(* IEC 61131-3 sources: Test-Git_ESME26/TestProgettoESME_26.fbsproj/AxisModuleLib Migration/DiagSource/AXM_FB_AxisModuleDiagSource.fb.st^, 38 files *)

(* ---- CancelWriting.meth.st ---- *)
{attribute 'conditionalshow_all_locals'}
METHOD INTERNAL CancelWriting : BOOL
VAR_INPUT
END_VAR

(* Deactivate writing if we are (for whatever reason) no longer adressed.
   May happen in case network connection with Diagnostics is disrupted or Source will be disabled *)

THIS^.diOldCmd			:= 0;
THIS^.diCmdExecState	:= 0;

(* ---- DiagQuit.meth.st ---- *)
{attribute 'conditionalshow_all_locals'}
METHOD INTERNAL DiagQuit : BOOL
VAR_INPUT
END_VAR

IF THIS^.i_xEnable AND THIS^.q_xActive AND THIS^.q_etDiag <> GD.ET_Diag.Ok AND THIS^.diState = 0 THEN

	THIS^.rtrigDiagQuit(CLK := THIS^.i_xDiagQuit);
	IF THIS^.rtrigDiagQuit.Q THEN
		CancelWriting();

		THIS^.udiOwnSourceId	:= 0;

		THIS^.fbTreeWriter.FB_Init(bInitRetains := FALSE, bInCopyCode := FALSE);

		THIS^.q_xReady		:= TRUE;
		THIS^.q_etDiag		:= GD.ET_Diag.Ok;
		THIS^.q_etDiagExt	:= AXM_ET_DiagExt.WaitUntilDiagnosticsManagerReady;
		THIS^.q_sMsg		:= '';

		THIS^.diState := 10;
	END_IF

END_IF

(* ---- ExceptionDuringWriting.meth.st ---- *)
{attribute 'conditionalshow_all_locals'}
METHOD INTERNAL ExceptionDuringWriting : BOOL
VAR_INPUT
END_VAR

(* exception during writing *)
CASE THIS^.etDiagExtTPL OF
	TPL.ET_DiagExt.TreeStartAlreadySuccessfullyCalled,
	TPL.ET_DiagExt.FileIdNotSet,
	TPL.ET_DiagExt.FileIdInvalid,
	TPL.ET_DiagExt.FileNotOpen,
	TPL.ET_DiagExt.UnexpectedFeedback,
	TPL.ET_DiagExt.TreeStartNotCalled,
	TPL.ET_DiagExt.TreeStartNotSuccessfullyCalled,
	TPL.ET_DiagExt.NoMoreNodeOpen,
	TPL.ET_DiagExt.CallTreeStartFirst,
	TPL.ET_DiagExt.NodesStillOpen:

		SetDiagOutputs(	i_etDiag	:= GD.ET_Diag.UnexpectedProgramBehavior,
						i_etDiagExt	:= AXM_ET_DiagExt.UnexpectedFeedback,
						i_sMsg		:= SE_CTBX.FC_MultiConcat(	i_sString1	:= 'FB_TreeWriter: ',
																i_sString2	:= GD.FC_EtDiagToString(THIS^.etDiag),
																i_sString3	:= ' - ',
																i_sString4	:= TPL.FC_EtDiagExtToString(THIS^.etDiagExtTPL)
															 )
					  );
	ELSE
		SetDiagOutputs(	i_etDiag	:= GD.ET_Diag.UnexpectedProgramBehavior,
						i_etDiagExt	:= AXM_ET_DiagExt.UnexpectedFeedback,
						i_sMsg		:= SE_CTBX.FC_MultiConcat(	i_sString1	:= 'FB_TreeWriter: ',
																i_sString2	:= GD.FC_EtDiagToString(THIS^.etDiag),
																i_sString3	:= ' - ',
																i_sString4	:= TPL.FC_EtDiagExtToString(THIS^.etDiagExtTPL)
															  )
					   );
END_CASE

CancelWriting();

(* ---- SetDiagOutputs.meth.st ---- *)
{attribute 'conditionalshow_all_locals'}
METHOD INTERNAL SetDiagOutputs : BOOL
VAR_INPUT
	i_etDiag		: GD.ET_Diag;
	i_etDiagExt		: AXM_ET_DiagExt;
	i_sMsg			: STRING[80];
END_VAR

IF THIS^.q_etDiag = GD.ET_Diag.Ok OR i_etDiagExt = AXM_ET_DiagExt.Disabled THEN

	IF i_etDiag <> GD.ET_Diag.Ok OR i_etDiagExt = AXM_ET_DiagExt.Disabled THEN

		IF i_etDiag <> GD.ET_Diag.Ok THEN
			THIS^.iq_stComStructure.iq_diCmd := -THIS^.iq_stComStructure.iq_diCmd;
		END_IF

		IF i_etDiagExt = AXM_ET_DiagExt.Disabled THEN
			THIS^.q_xActive := FALSE;

			CancelWriting();
		END_IF

		THIS^.q_xReady := FALSE;
		THIS^.diState := 0;
	END_IF

	THIS^.q_etDiag		:= i_etDiag;
	THIS^.q_etDiagExt	:= i_etDiagExt;
	THIS^.q_sMsg		:= i_sMsg;

END_IF

(* ---- WriteDiagDataControl.meth.st ---- *)
{attribute 'conditionalshow_all_locals'}
METHOD INTERNAL WriteDiagDataControl : BOOL
VAR_INPUT
END_VAR

IF (THIS^.diOldCmd <> THIS^.iq_stComStructure.iq_diCmd AND THIS^.iq_stComStructure.iq_diCmd > 0) THEN

	THIS^.diOldCmd := THIS^.iq_stComStructure.iq_diCmd;

	(* new command, start execution *)
	CASE THIS^.iq_stComStructure.iq_diCmd OF

		1: (* write diag data to file *)
			IF (THIS^.iq_stComStructure.i_diFileId > 0) THEN

				SetDiagOutputs(	i_etDiag		:= GD.ET_Diag.Ok,
								i_etDiagExt		:= AXM_ET_DiagExt.WritingToFile,
								i_sMsg			:= '');

				THIS^.iq_stComStructure.q_lrProgress := 0.0;

				THIS^.fbTreeWriter.diFileId := THIS^.iq_stComStructure.i_diFileId;

				THIS^.diCmdExecState := 1; (* start writing to file *)
			ELSE
				(* invalid file id *)
				SetDiagOutputs(	i_etDiag		:= GD.ET_Diag.InputParameterInvalid,
								i_etDiagExt		:= AXM_ET_DiagExt.FileIdInvalid,
								i_sMsg			:= CONCAT('Invalid file Id iq_stComStructure.i_diFileId: ', TO_STRING(THIS^.iq_stComStructure.i_diFileId)));
			END_IF
		ELSE
			(* unkown cmd *)
			SetDiagOutputs(	i_etDiag		:= GD.ET_Diag.InputParameterInvalid,
							i_etDiagExt		:= AXM_ET_DiagExt.CmdUnknown,
							i_sMsg			:= CONCAT('Unknown command iq_stComStructure.diCmd: ', DINT_TO_STRING(THIS^.iq_stComStructure.iq_diCmd)));

			CancelWriting();
	END_CASE
END_IF

(* ---- WriteDiagDataToFile.meth.st ---- *)
{attribute 'conditionalshow_all_locals'}
METHOD INTERNAL WriteDiagDataToFile : BOOL
VAR_INPUT
END_VAR
VAR
END_VAR

TPL.FC_CanContinueWriting(iq_stCanContinueWriting := THIS^.iq_stComStructure.iq_stCanContinueWriting); (* loop as long as we can continue to write *)

WHILE (THIS^.iq_stComStructure.iq_stCanContinueWriting.xCanContinue) DO

	CASE THIS^.diCmdExecState OF
		1:
			THIS^.pstTmp := ADR(THIS^.iq_stMachineItf);

			(* start writing *)
			THIS^.fbTreeWriter.TreeStart(	i_sName					:= THIS^.c_sName,
											i_sTypeName				:= THIS^.c_sTypeName,
											i_sTitleEnglish			:= 'AxisModule interface',
											i_sTitleGerman			:= 'AxisModule Schnittstelle',
											i_uiPrintRank			:= 14,
											i_sEmptyListTextEnglish	:= 'No data available to show',
											i_sEmptyListTextGerman	:= 'Keine Daten zum Anzeigen vorhanden',
											q_etDiag				=> THIS^.etDiag,
											q_etDiagExt				=> THIS^.etDiagExtTPL,
											q_sMsg					=> THIS^.sMsg);

			IF THIS^.etDiag <> GD.ET_Diag.Ok THEN
				ExceptionDuringWriting();
				EXIT;
			END_IF

			THIS^.audiHierarchy[1]	:= 1;
			THIS^.apstHierarchy[1]	:= THIS^.pstTmp;
			THIS^.udiLevelCounter	:= 1; (* start loop at index 1 *)

			THIS^.diCmdExecState := THIS^.diCmdExecState + 1;

        2:
			(* writing node main machine *)
			THIS^.sModuleName := CONCAT(UDINT_TO_STRING(THIS^.pstTmp^.i_udiModuleId), ' : ');
			THIS^.sModuleName := CONCAT(THIS^.sModuleName, THIS^.pstTmp^.i_sModuleName);

			THIS^.fbTreeWriter.NodeStart(	i_sName		:= THIS^.sModuleName,
											q_etDiag	=> THIS^.etDiag,
											q_etDiagExt	=> THIS^.etDiagExtTPL,
											q_sMsg		=> THIS^.sMsg);

			IF THIS^.etDiag <> GD.ET_Diag.Ok THEN
				ExceptionDuringWriting();
				EXIT;
			END_IF

			IF (THIS^.pstTmp^.iq_stExt.udiNumberOfSubModules <> 0) THEN
				THIS^.diCmdExecState := THIS^.diCmdExecState + 1;
			ELSE
				THIS^.fbTreeWriter.NodeEnd(	q_etDiag	=> THIS^.etDiag,
											q_etDiagExt	=> THIS^.etDiagExtTPL,
											q_sMsg		=> THIS^.sMsg);

				IF THIS^.etDiag <> GD.ET_Diag.Ok THEN
					ExceptionDuringWriting();
					EXIT;
				END_IF

				THIS^.diCmdExecState := 4;
			END_IF

		3:
			(* Navigate to next module *)
			(* Try to go down *)
			IF ((THIS^.apstHierarchy[THIS^.udiLevelCounter]^.iq_stExt.udiNumberOfSubModules > 0) AND (THIS^.udiLevelCounter < THIS^.c_udiMaxLevel)) THEN
				(* Go down *)
				THIS^.udiLevelCounter := THIS^.udiLevelCounter + 1;
				THIS^.audiHierarchy[THIS^.udiLevelCounter] := 1;
				(* Set pointer *)
				THIS^.apstHierarchy[THIS^.udiLevelCounter] := THIS^.apstHierarchy[THIS^.udiLevelCounter - 1]^.iq_stExt.dwSubModulesItf
					+ UDINT_TO_DWORD((THIS^.audiHierarchy[THIS^.udiLevelCounter] - 1) * SIZEOF(THIS^.pstTmp^));

			ELSIF (THIS^.apstHierarchy[THIS^.udiLevelCounter - 1] <> 0) THEN
				(* Cannot go down *)

				(* Write end-tag of last module *)
				THIS^.fbTreeWriter.NodeEnd(	q_etDiag	=> THIS^.etDiag,
											q_etDiagExt	=> THIS^.etDiagExtTPL,
											q_sMsg		=> THIS^.sMsg);

				IF THIS^.etDiag <> GD.ET_Diag.Ok THEN
					ExceptionDuringWriting();
					EXIT;
				END_IF

				(* Check if you can go right *)
				IF (THIS^.apstHierarchy[THIS^.udiLevelCounter - 1]^.iq_stExt.udiNumberOfSubModules > THIS^.audiHierarchy[THIS^.udiLevelCounter]) THEN
					(* Go right *)
					THIS^.audiHierarchy[THIS^.udiLevelCounter] := THIS^.audiHierarchy[THIS^.udiLevelCounter] + 1;
					(* Set pointer *)
					THIS^.apstHierarchy[THIS^.udiLevelCounter] := THIS^.apstHierarchy[THIS^.udiLevelCounter - 1]^.iq_stExt.dwSubModulesItf
						+  UDINT_TO_DWORD((THIS^.audiHierarchy[THIS^.udiLevelCounter] - 1) * SIZEOF(THIS^.pstTmp^));
				ELSE
					(* Check if you can go up *)
					(* Go up until you can go right *)
					THIS^.xLoop := TRUE;
					WHILE (THIS^.xLoop AND (THIS^.udiLevelCounter > 1)) DO
						THIS^.udiLevelCounter := THIS^.udiLevelCounter - 1;
						IF (THIS^.udiLevelCounter > 1) THEN
							THIS^.xLoop := (THIS^.apstHierarchy[THIS^.udiLevelCounter - 1]^.iq_stExt.udiNumberOfSubModules <= THIS^.audiHierarchy[THIS^.udiLevelCounter]);
							IF (THIS^.xLoop) THEN
								(* Write end-tag of last module *)
				  				THIS^.fbTreeWriter.NodeEnd(	q_etDiag	=> THIS^.etDiag,
															q_etDiagExt	=> THIS^.etDiagExtTPL,
															q_sMsg		=> THIS^.sMsg);

								IF THIS^.etDiag <> GD.ET_Diag.Ok THEN
									ExceptionDuringWriting();
									EXIT;
								END_IF
							END_IF
						ELSE
							THIS^.xLoop := FALSE;
						END_IF
					END_WHILE

					(* Write end-tag of last module *)
					THIS^.fbTreeWriter.NodeEnd(	q_etDiag	=> THIS^.etDiag,
												q_etDiagExt	=> THIS^.etDiagExtTPL,
												q_sMsg		=> THIS^.sMsg);

					IF THIS^.etDiag <> GD.ET_Diag.Ok THEN
						ExceptionDuringWriting();
						EXIT;
					END_IF

					IF (THIS^.udiLevelCounter <= 1) THEN
						(* End of tree reached *)
						THIS^.diCmdExecState := 4;
					ELSE
						(* Go right *)
						(* Set pointer *)
						THIS^.audiHierarchy[THIS^.udiLevelCounter] := THIS^.audiHierarchy[THIS^.udiLevelCounter] + 1;
						THIS^.apstHierarchy[THIS^.udiLevelCounter] := THIS^.apstHierarchy[THIS^.udiLevelCounter - 1]^.iq_stExt.dwSubModulesItf
							+  UDINT_TO_DWORD((THIS^.audiHierarchy[THIS^.udiLevelCounter] - 1) * SIZEOF(THIS^.pstTmp^));
					END_IF
				END_IF
			END_IF

			(* Write node of current module *)
			IF (THIS^.diCmdExecState <> 4) THEN
				IF (THIS^.apstHierarchy[THIS^.udiLevelCounter] <> 0) THEN
					(* Set name pointer to character before last semicolon *)
					THIS^.pstChar := ADR(THIS^.apstHierarchy[THIS^.udiLevelCounter]^.i_sModuleName) +  INT_TO_DWORD((LEN(THIS^.apstHierarchy[THIS^.udiLevelCounter]^.i_sModuleName) - 3));
					THIS^.sModuleName := THIS^.pstChar^;
					(* Search for beginning of module name *)
					WHILE (FIND(THIS^.sModuleName, ':') <> 1) DO
						THIS^.pstChar := THIS^.pstChar - 1;
						THIS^.sModuleName := THIS^.pstChar^;
					END_WHILE
					(* Make string nicer *)
					THIS^.sModuleName := CONCAT (' ', THIS^.sModuleName);

					THIS^.fbTreeWriter.NodeStart(	i_sName		:= CONCAT(UDINT_TO_STRING(THIS^.apstHierarchy[THIS^.udiLevelCounter]^.i_udiModuleId), THIS^.sModuleName),
													q_etDiag	=> THIS^.etDiag,
													q_etDiagExt	=> THIS^.etDiagExtTPL,
													q_sMsg		=> THIS^.sMsg);

					IF THIS^.etDiag <> GD.ET_Diag.Ok THEN
						ExceptionDuringWriting();
						EXIT;
					END_IF

					(* is an axis module? *)
					IF (THIS^.apstHierarchy[THIS^.udiLevelCounter]^.q_dwModuleType =  UDINT_TO_DWORD(TPL.ET_ModuleType.AxisModule)) THEN
						IF (THIS^.apstHierarchy[THIS^.udiLevelCounter]^.q_udiModuleVersion <> 1) THEN
							(* version not supported *)
							THIS^.fbTreeWriter.Parameter(	i_sName		:= 'Exception',
															i_sValue	:= 'Version of AxisModule not supported',
															q_etDiag	=> THIS^.etDiag,
															q_etDiagExt	=> THIS^.etDiagExtTPL,
															q_sMsg		=> THIS^.sMsg);

							IF THIS^.etDiag <> GD.ET_Diag.Ok THEN
								ExceptionDuringWriting();
								EXIT;
							END_IF
						ELSE
							(* print additional interface *)
							THIS^.pstInterface := 0;
							(* get pointer to additional interface *)
							IF (THIS^.udiLevelCounter >= 2) THEN
								IF(THIS^.apstHierarchy[THIS^.udiLevelCounter - 1] <> 0) THEN
									IF (THIS^.apstHierarchy[THIS^.udiLevelCounter - 1]^.iq_stExt.pdwSubModulesAddItf <> 0) THEN
										(* get correct position in list of add interface pointers *)
										THIS^.pdw := THIS^.apstHierarchy[THIS^.udiLevelCounter - 1]^.iq_stExt.pdwSubModulesAddItf
											+ UDINT_TO_DWORD((THIS^.audiHierarchy[THIS^.udiLevelCounter](* number OF submodule *) - 1) * SIZEOF(THIS^.pdw^));
										IF (THIS^.pdw^ <> 0) THEN
											THIS^.pstInterface := THIS^.pdw^;
										END_IF
									END_IF
								END_IF
							END_IF

							IF (THIS^.pstInterface = 0) THEN
								THIS^.fbTreeWriter.Parameter(	i_sName		:= 'Exception',
																i_sValue	:= 'Could not get pointer to additional interface',
																q_etDiag	=> THIS^.etDiag,
																q_etDiagExt	=> THIS^.etDiagExtTPL,
																q_sMsg		=> THIS^.sMsg);

								IF THIS^.etDiag <> GD.ET_Diag.Ok THEN
									ExceptionDuringWriting();
									EXIT;
								END_IF
							ELSE
								THIS^.diCmdExecState := 5; (* continue output in different state *)
							END_IF (* addinterface pointer *)
						END_IF (* version *)
					END_IF (* module type *)
				END_IF
			END_IF

		4:
			(* library versions *)
			THIS^.fbTreeWriter.NodeStart(	i_sName		:= 'LibraryVersions',
											q_etDiag	=> THIS^.etDiag,
											q_etDiagExt	=> THIS^.etDiagExtTPL,
											q_sMsg		=> THIS^.sMsg);

			IF THIS^.etDiag <> GD.ET_Diag.Ok THEN
				ExceptionDuringWriting();
				EXIT;
			END_IF

				THIS^.fbTreeWriter.Parameter(	i_sName		:= 'GlobalDiagnostics',
												i_sValue	:= GD.Gc_sLibraryVersion,
												q_etDiag	=> THIS^.etDiag,
												q_etDiagExt	=> THIS^.etDiagExtTPL,
												q_sMsg		=> THIS^.sMsg);

				IF THIS^.etDiag <> GD.ET_Diag.Ok THEN
					ExceptionDuringWriting();
					EXIT;
				END_IF

				THIS^.fbTreeWriter.Parameter(	i_sName		:= 'PLCopenMcPart1',
												i_sValue	:= 'TODO', //PLCO. PDL_Gc_sLibraryVersion,
												q_etDiag	=> THIS^.etDiag,
												q_etDiagExt	=> THIS^.etDiagExtTPL,
												q_sMsg		=> THIS^.sMsg);

				IF THIS^.etDiag <> GD.ET_Diag.Ok THEN
					ExceptionDuringWriting();
					EXIT;
				END_IF

			THIS^.fbTreeWriter.NodeEnd(	q_etDiag	=> THIS^.etDiag,
										q_etDiagExt	=> THIS^.etDiagExtTPL,
										q_sMsg		=> THIS^.sMsg);

			IF THIS^.etDiag <> GD.ET_Diag.Ok THEN
				ExceptionDuringWriting();
				EXIT;
			END_IF

			THIS^.fbTreeWriter.TreeEnd(	q_etDiag	=> THIS^.etDiag,
										q_etDiagExt	=> THIS^.etDiagExtTPL,
										q_sMsg		=> THIS^.sMsg);

			IF THIS^.etDiag <> GD.ET_Diag.Ok THEN
				ExceptionDuringWriting();
				EXIT;
			END_IF
			(* done *)

			(* signal command execution *)
			THIS^.iq_stComStructure.iq_diCmd := 0;

			SetDiagOutputs(	i_etDiag	:= GD.ET_Diag.Ok,
							i_etDiagExt	:= AXM_ET_DiagExt.DataSuccessfullyWritten,
							i_sMsg		:= '');

			THIS^.diCmdExecState := 0;
			EXIT; (* exit the while loop *)

		5:
			(* continue output of AxisModule interface *)
			WriteInterfaceStart(q_etDiag	=> THIS^.etDiag,
								q_etDiagExt	=> THIS^.etDiagExtTPL,
								q_sMsg		=> THIS^.sMsg);

			IF THIS^.etDiag <> GD.ET_Diag.Ok THEN
				ExceptionDuringWriting();
				EXIT;
			END_IF

			THIS^.diCmdExecState := 51;

		51:
			WriteInterfaceMain(	q_etDiag	=> THIS^.etDiag,
								q_etDiagExt	=> THIS^.etDiagExtTPL,
								q_sMsg		=> THIS^.sMsg);

			IF THIS^.etDiag <> GD.ET_Diag.Ok THEN
				ExceptionDuringWriting();
				EXIT;
			END_IF

			THIS^.diCmdExecState := 52;

		52:
			WriteInterfaceHomeStart(q_etDiag	=> THIS^.etDiag,
									q_etDiagExt	=> THIS^.etDiagExtTPL,
									q_sMsg		=> THIS^.sMsg);

			IF THIS^.etDiag <> GD.ET_Diag.Ok THEN
				ExceptionDuringWriting();
				EXIT;
			END_IF

			THIS^.diCmdExecState := 53;

		53:
			WriteInterfaceHomeParam(q_etDiag	=> THIS^.etDiag,
									q_etDiagExt	=> THIS^.etDiagExtTPL,
									q_sMsg		=> THIS^.sMsg);

			IF THIS^.etDiag <> GD.ET_Diag.Ok THEN
				ExceptionDuringWriting();
				EXIT;
			END_IF

			THIS^.diCmdExecState := 54;

		54:
// 			WriteInterfaceHomeTouchProbe(	q_etDiag	=> THIS^.etDiag,
// 											q_etDiagExt	=> THIS^.etDiagExtTPL,
// 											q_sMsg		=> THIS^.sMsg);
//
// 			IF THIS^.etDiag <> GD.ET_Diag.Ok THEN
// 				ExceptionDuringWriting();
// 				EXIT;
// 			END_IF

			THIS^.diCmdExecState := 55;

		55:
// 			WriteInterfaceHomeSensor(	q_etDiag	=> THIS^.etDiag,
// 										q_etDiagExt	=> THIS^.etDiagExtTPL,
// 										q_sMsg		=> THIS^.sMsg);
// 			WriteInterfaceHomeDigitalInput(	q_etDiag	=> THIS^.etDiag,
// 											q_etDiagExt	=> THIS^.etDiagExtTPL,
// 											q_sMsg		=> THIS^.sMsg);
//
// 			IF THIS^.etDiag <> GD.ET_Diag.Ok THEN
// 				ExceptionDuringWriting();
// 				EXIT;
// 			END_IF

			THIS^.diCmdExecState := 56;

		56:
// 			WriteInterfaceHomeLimitSwitch(	q_etDiag	=> THIS^.etDiag,
// 											q_etDiagExt	=> THIS^.etDiagExtTPL,
// 											q_sMsg		=> THIS^.sMsg);
//
// 			IF THIS^.etDiag <> GD.ET_Diag.Ok THEN
// 				ExceptionDuringWriting();
// 				EXIT;
// 			END_IF

			THIS^.diCmdExecState := 57;

		57:
// 			WriteInterfaceHomeTorque(	q_etDiag	=> THIS^.etDiag,
// 										q_etDiagExt	=> THIS^.etDiagExtTPL,
// 										q_sMsg		=> THIS^.sMsg);
//
// 			IF THIS^.etDiag <> GD.ET_Diag.Ok THEN
// 				ExceptionDuringWriting();
// 				EXIT;
// 			END_IF

			THIS^.diCmdExecState := 581;

		581:
// 			WriteInterfaceHomeForce(	q_etDiag	=> THIS^.etDiag,
// 										q_etDiagExt	=> THIS^.etDiagExtTPL,
// 										q_sMsg		=> THIS^.sMsg);
//
// 			IF THIS^.etDiag <> GD.ET_Diag.Ok THEN
// 				ExceptionDuringWriting();
// 				EXIT;
// 			END_IF

			THIS^.diCmdExecState := 58;

		58:
			WriteInterfaceHomeMoveOnPos(q_etDiag	=> THIS^.etDiag,
										q_etDiagExt	=> THIS^.etDiagExtTPL,
										q_sMsg		=> THIS^.sMsg);

			IF THIS^.etDiag <> GD.ET_Diag.Ok THEN
				ExceptionDuringWriting();
				EXIT;
			END_IF

			THIS^.diCmdExecState := 59;

		59:
			WriteInterfaceHomeSetPos(	q_etDiag	=> THIS^.etDiag,
										q_etDiagExt	=> THIS^.etDiagExtTPL,
										q_sMsg		=> THIS^.sMsg);

			IF THIS^.etDiag <> GD.ET_Diag.Ok THEN
				ExceptionDuringWriting();
				EXIT;
			END_IF

			THIS^.diCmdExecState := 60;

		60:
// 			WriteInterfaceHomeWritePos(	q_etDiag	=> THIS^.etDiag,
// 										q_etDiagExt	=> THIS^.etDiagExtTPL,
// 										q_sMsg		=> THIS^.sMsg);
//
// 			IF THIS^.etDiag <> GD.ET_Diag.Ok THEN
// 				ExceptionDuringWriting();
// 				EXIT;
// 			END_IF

			THIS^.diCmdExecState := 61;

		61:
			WriteInterfaceHomeEnd(	q_etDiag	=> THIS^.etDiag,
									q_etDiagExt	=> THIS^.etDiagExtTPL,
									q_sMsg		=> THIS^.sMsg);

			IF THIS^.etDiag <> GD.ET_Diag.Ok THEN
				ExceptionDuringWriting();
				EXIT;
			END_IF

			THIS^.diCmdExecState := 62;

		62:
			WriteInterfaceManual(	q_etDiag	=> THIS^.etDiag,
									q_etDiagExt	=> THIS^.etDiagExtTPL,
									q_sMsg		=> THIS^.sMsg);

			IF THIS^.etDiag <> GD.ET_Diag.Ok THEN
				ExceptionDuringWriting();
				EXIT;
			END_IF

			THIS^.diCmdExecState := 63;

		63:
			WriteInterfaceEndless(	q_etDiag	=> THIS^.etDiag,
									q_etDiagExt	=> THIS^.etDiagExtTPL,
									q_sMsg		=> THIS^.sMsg);

			IF THIS^.etDiag <> GD.ET_Diag.Ok THEN
				ExceptionDuringWriting();
				EXIT;
			END_IF

			THIS^.diCmdExecState := 64;

		64:
			WriteInterfaceMultiCamStart(q_etDiag	=> THIS^.etDiag,
										q_etDiagExt	=> THIS^.etDiagExtTPL,
										q_sMsg		=> THIS^.sMsg);

			IF THIS^.etDiag <> GD.ET_Diag.Ok THEN
				ExceptionDuringWriting();
				EXIT;
			END_IF

			THIS^.diCmdExecState := 65;

		65:
			WriteInterfaceMultiCamParamIn(	q_etDiag	=> THIS^.etDiag,
											q_etDiagExt	=> THIS^.etDiagExtTPL,
											q_sMsg		=> THIS^.sMsg);

			IF THIS^.etDiag <> GD.ET_Diag.Ok THEN
				ExceptionDuringWriting();
				EXIT;
			END_IF

			THIS^.diCmdExecState := 66;

		66:
			WriteInterfaceMultiCamMotionParStart(	q_etDiag	=> THIS^.etDiag,
													q_etDiagExt	=> THIS^.etDiagExtTPL,
													q_sMsg		=> THIS^.sMsg);

			IF THIS^.etDiag <> GD.ET_Diag.Ok THEN
				ExceptionDuringWriting();
				EXIT;
			END_IF

			(* loop over multiple cycles in state 67 and 68 *)
			(* FOR diMotionParCounter := 0 TO Gc_udiMaxNumberOfCamTables DO *)
			THIS^.diMotionParCounter := -1;

			THIS^.diCmdExecState := 67;

		67:
			IF (THIS^.i_xPrintCamData) THEN (* allow the user to protect his know-how *)
				IF (THIS^.diMotionParCounter < UDINT_TO_DINT(AXM_GPL.Gc_udiMaxNumberOfCamTables)) THEN (* loop over more than one cycle *)

					THIS^.diMotionParCounter := THIS^.diMotionParCounter + 1;

					WriteInterfaceMultiCamMotionParCyclicStart(	q_etDiag	=> THIS^.etDiag,
																q_etDiagExt	=> THIS^.etDiagExtTPL,
																q_sMsg		=> THIS^.sMsg);
					(* loop over multiple cycles in state 553 *)
					(* FOR diCamPointerCounter := 0 TO MAX_NO_OF_SEG DO *)
					THIS^.diCamPointCounter := 0;
					THIS^.diCmdExecState := 1000; (* switch to loop over CamPoints *)
				ELSE
					THIS^.diCmdExecState := 999;
				END_IF
			ELSE
				THIS^.fbTreeWriter.Parameter(	i_sName		:= 'data omitted',
												i_sValue	:= 'because i_xPrintCamData is FALSE',
												q_etDiag	=> THIS^.etDiag,
												q_etDiagExt	=> THIS^.etDiagExtTPL,
												q_sMsg		=> THIS^.sMsg);

				IF THIS^.etDiag <> GD.ET_Diag.Ok THEN
					ExceptionDuringWriting();
					EXIT;
				END_IF

				diCmdExecState := 999;
			END_IF

		1000:
			WriteInterfaceMultiCamMotionParCamPointStart(	q_etDiag	=> THIS^.etDiag,
															q_etDiagExt	=> THIS^.etDiagExtTPL,
															q_sMsg		=> THIS^.sMsg);

			IF THIS^.etDiag <> GD.ET_Diag.Ok THEN
				ExceptionDuringWriting();
				EXIT;
			END_IF

			THIS^.diCmdExecState := 68;

		68: (* loop over cam points using diCamPointerCounter *)
			IF (THIS^.diCamPointCounter <= 32) THEN

				WriteInterfaceMultiCamMotionParCamPoint(q_etDiag	=> THIS^.etDiag,
														q_etDiagExt	=> THIS^.etDiagExtTPL,
														q_sMsg		=> THIS^.sMsg);

				IF THIS^.etDiag <> GD.ET_Diag.Ok THEN
					ExceptionDuringWriting();
					EXIT;
				END_IF

				THIS^.diCamPointCounter := THIS^.diCamPointCounter + 1;
			ELSE
				WriteInterfaceMultiCamMotionParCamPointEnd(	q_etDiag	=> THIS^.etDiag,
															q_etDiagExt	=> THIS^.etDiagExtTPL,
															q_sMsg		=> THIS^.sMsg);

				IF THIS^.etDiag <> GD.ET_Diag.Ok THEN
					ExceptionDuringWriting();
					EXIT;
				END_IF

				THIS^.diCmdExecState := 1001;
			END_IF

		1001:
				WriteInterfaceMultiCamMotionParCyclicEnd(	q_etDiag	=> THIS^.etDiag,
															q_etDiagExt	=> THIS^.etDiagExtTPL,
															q_sMsg		=> THIS^.sMsg);

				IF THIS^.etDiag <> GD.ET_Diag.Ok THEN
					ExceptionDuringWriting();
					EXIT;
				END_IF

				THIS^.diCmdExecState := 67;
		999:
			WriteInterfaceMultiCamMotionParEnd(	q_etDiag	=> THIS^.etDiag,
												q_etDiagExt	=> THIS^.etDiagExtTPL,
												q_sMsg		=> THIS^.sMsg);

			IF THIS^.etDiag <> GD.ET_Diag.Ok THEN
				ExceptionDuringWriting();
				EXIT;
			END_IF

			THIS^.diCmdExecState := 70;

		70:
			WriteInterfaceMultiCamExt(	q_etDiag	=> THIS^.etDiag,
										q_etDiagExt	=> THIS^.etDiagExtTPL,
										q_sMsg		=> THIS^.sMsg);

			IF THIS^.etDiag <> GD.ET_Diag.Ok THEN
				ExceptionDuringWriting();
				EXIT;
			END_IF

			THIS^.diCmdExecState := 71;

		71:
			WriteInterfaceMultiCamParamOut(	q_etDiag	=> THIS^.etDiag,
											q_etDiagExt	=> THIS^.etDiagExtTPL,
											q_sMsg		=> THIS^.sMsg);

			IF THIS^.etDiag <> GD.ET_Diag.Ok THEN
				ExceptionDuringWriting();
				EXIT;
			END_IF

			THIS^.diCmdExecState := 72;

		72:
			WriteInterfaceMultiCamParamOutActualCamData(	q_etDiag	=> THIS^.etDiag,
															q_etDiagExt	=> THIS^.etDiagExtTPL,
															q_sMsg		=> THIS^.sMsg);

			IF THIS^.etDiag <> GD.ET_Diag.Ok THEN
				ExceptionDuringWriting();
				EXIT;
			END_IF

			THIS^.diCmdExecState := 73;

		73:
			WriteInterfaceMultiCamEnd(	q_etDiag	=> THIS^.etDiag,
										q_etDiagExt	=> THIS^.etDiagExtTPL,
										q_sMsg		=> THIS^.sMsg);

			IF THIS^.etDiag <> GD.ET_Diag.Ok THEN
				ExceptionDuringWriting();
				EXIT;
			END_IF

			THIS^.diCmdExecState := 74;

		74:
			WriteInterfacePos(	q_etDiag	=> THIS^.etDiag,
								q_etDiagExt	=> THIS^.etDiagExtTPL,
								q_sMsg		=> THIS^.sMsg);

			IF THIS^.etDiag <> GD.ET_Diag.Ok THEN
				ExceptionDuringWriting();
				EXIT;
			END_IF

			THIS^.diCmdExecState := 75;

		75:
			WriteInterfaceBrake(q_etDiag	=> THIS^.etDiag,
								q_etDiagExt	=> THIS^.etDiagExtTPL,
								q_sMsg		=> THIS^.sMsg);

			IF THIS^.etDiag <> GD.ET_Diag.Ok THEN
				ExceptionDuringWriting();
				EXIT;
			END_IF

			THIS^.diCmdExecState := 76;

		76:
			WriteInterfaceAdditionalMode(	q_etDiag	=> THIS^.etDiag,
											q_etDiagExt	=> THIS^.etDiagExtTPL,
											q_sMsg		=> THIS^.sMsg);

			IF THIS^.etDiag <> GD.ET_Diag.Ok THEN
				ExceptionDuringWriting();
				EXIT;
			END_IF

			THIS^.diCmdExecState := 77;

		77:

			WriteInterfaceEnd(	q_etDiag	=> THIS^.etDiag,
								q_etDiagExt	=> THIS^.etDiagExtTPL,
								q_sMsg		=> THIS^.sMsg);

			IF THIS^.etDiag <> GD.ET_Diag.Ok THEN
				ExceptionDuringWriting();
				EXIT;
			END_IF

			THIS^.diCmdExecState := 3; (* go to next module *)

	END_CASE

	(* check again whether we can continue writing *)
	TPL.FC_CanContinueWriting(iq_stCanContinueWriting := THIS^.iq_stComStructure.iq_stCanContinueWriting);
END_WHILE

(* ---- WriteInterfaceAdditionalMode.meth.st ---- *)
{attribute 'conditionalshow_all_locals'}
METHOD INTERNAL WriteInterfaceAdditionalMode : BOOL
VAR_INPUT
END_VAR
VAR_OUTPUT
	q_etDiag		: GD.ET_Diag;
	q_etDiagExt	: TPL.ET_DiagExt;
	q_sMsg			: STRING[80];
END_VAR

THIS^.fbTreeWriter.NodeStart(	i_sName		:= 'stAdditional',
								q_etDiag	=> q_etDiag,
								q_etDiagExt	=> q_etDiagExt,
								q_sMsg		=> q_sMsg);

IF q_etDiag <> GD.ET_Diag.Ok THEN
	RETURN;
END_IF

	THIS^.fbTreeWriter.Parameter(	i_sName		:= 'i_etDiag',
									i_sValue	:= GD.FC_EtDiagToString(THIS^.pstInterface^.stAdditional.i_etDiag),
									q_etDiag	=> q_etDiag,
									q_etDiagExt	=> q_etDiagExt,
									q_sMsg		=> q_sMsg);

	IF q_etDiag <> GD.ET_Diag.Ok THEN
		RETURN;
	END_IF

	THIS^.fbTreeWriter.Parameter(	i_sName		:= 'i_udiDiagExt',
									i_sValue	:= UDINT_TO_STRING(THIS^.pstInterface^.stAdditional.i_udiDiagExt),
									q_etDiag	=> q_etDiag,
									q_etDiagExt	=> q_etDiagExt,
									q_sMsg		=> q_sMsg);

	IF q_etDiag <> GD.ET_Diag.Ok THEN
		RETURN;
	END_IF

	THIS^.fbTreeWriter.Parameter(	i_sName		:= 'i_sDiagExt',
									i_sValue	:= THIS^.pstInterface^.stAdditional.i_sDiagExt,
									q_etDiag	=> q_etDiag,
									q_etDiagExt	=> q_etDiagExt,
									q_sMsg		=> q_sMsg);

	IF q_etDiag <> GD.ET_Diag.Ok THEN
		RETURN;
	END_IF

	THIS^.fbTreeWriter.Parameter(	i_sName		:= 'i_sMsg',
									i_sValue	:= THIS^.pstInterface^.stAdditional.i_sMsg,
									q_etDiag	=> q_etDiag,
									q_etDiagExt	=> q_etDiagExt,
									q_sMsg		=> q_sMsg);

	IF q_etDiag <> GD.ET_Diag.Ok THEN
		RETURN;
	END_IF

	THIS^.fbTreeWriter.Parameter(	i_sName		:= 'i_xActive',
									i_sValue	:= BOOL_TO_STRING(THIS^.pstInterface^.stAdditional.i_xActive),
									q_etDiag	=> q_etDiag,
									q_etDiagExt	=> q_etDiagExt,
									q_sMsg		=> q_sMsg);

	IF q_etDiag <> GD.ET_Diag.Ok THEN
		RETURN;
	END_IF

	THIS^.fbTreeWriter.Parameter(	i_sName		:= 'i_xReady',
									i_sValue	:= BOOL_TO_STRING(THIS^.pstInterface^.stAdditional.i_xReady),
									q_etDiag	=> q_etDiag,
									q_etDiagExt	=> q_etDiagExt,
									q_sMsg		=> q_sMsg);

	IF q_etDiag <> GD.ET_Diag.Ok THEN
		RETURN;
	END_IF

	THIS^.fbTreeWriter.Parameter(	i_sName		:= 'i_xActionCmdDone',
									i_sValue	:= BOOL_TO_STRING(THIS^.pstInterface^.stAdditional.i_xActionCmdDone),
									q_etDiag	=> q_etDiag,
									q_etDiagExt	=> q_etDiagExt,
									q_sMsg		=> q_sMsg);

	IF q_etDiag <> GD.ET_Diag.Ok THEN
		RETURN;
	END_IF

	THIS^.fbTreeWriter.Parameter(	i_sName		:= 'q_xEnable',
									i_sValue	:= BOOL_TO_STRING(THIS^.pstInterface^.stAdditional.q_xEnable),
									q_etDiag	=> q_etDiag,
									q_etDiagExt	=> q_etDiagExt,
									q_sMsg		=> q_sMsg);

	IF q_etDiag <> GD.ET_Diag.Ok THEN
		RETURN;
	END_IF

	THIS^.fbTreeWriter.Parameter(	i_sName		:= 'q_xStart',
									i_sValue	:= BOOL_TO_STRING(THIS^.pstInterface^.stAdditional.q_xStart),
									q_etDiag	=> q_etDiag,
									q_etDiagExt	=> q_etDiagExt,
									q_sMsg		=> q_sMsg);

	IF q_etDiag <> GD.ET_Diag.Ok THEN
		RETURN;
	END_IF

	THIS^.fbTreeWriter.Parameter(	i_sName		:= 'q_xWsSelect',
									i_sValue	:= BOOL_TO_STRING(THIS^.pstInterface^.stAdditional.q_xWsSelect),
									q_etDiag	=> q_etDiag,
									q_etDiagExt	=> q_etDiagExt,
									q_sMsg		=> q_sMsg);

	IF q_etDiag <> GD.ET_Diag.Ok THEN
		RETURN;
	END_IF

	THIS^.fbTreeWriter.Parameter(	i_sName		:= 'q_xWsStart',
									i_sValue	:= BOOL_TO_STRING(THIS^.pstInterface^.stAdditional.q_xWsStart),
									q_etDiag	=> q_etDiag,
									q_etDiagExt	=> q_etDiagExt,
									q_sMsg		=> q_sMsg);

	IF q_etDiag <> GD.ET_Diag.Ok THEN
		RETURN;
	END_IF

THIS^.fbTreeWriter.NodeEnd(	q_etDiag	=> q_etDiag,
							q_etDiagExt	=> q_etDiagExt,
							q_sMsg		=> q_sMsg);

IF q_etDiag <> GD.ET_Diag.Ok THEN
	RETURN;
END_IF

(* ---- WriteInterfaceBrake.meth.st ---- *)
{attribute 'conditionalshow_all_locals'}
METHOD INTERNAL WriteInterfaceBrake : BOOL
VAR_INPUT
END_VAR
VAR_OUTPUT
	q_etDiag		: GD.ET_Diag;
	q_etDiagExt	: TPL.ET_DiagExt;
	q_sMsg			: STRING[80];
END_VAR

THIS^.fbTreeWriter.NodeStart(	i_sName		:= 'stBrake',
								q_etDiag	=> q_etDiag,
								q_etDiagExt	=> q_etDiagExt,
								q_sMsg		=> q_sMsg);

IF q_etDiag <> GD.ET_Diag.Ok THEN
	RETURN;
END_IF

	THIS^.fbTreeWriter.Parameter(	i_sName		:= 'q_xBrakeReleased',
									i_sValue	:= BOOL_TO_STRING(THIS^.pstInterface^.stBrake.q_xBrakeReleased),
									q_etDiag	=> q_etDiag,
									q_etDiagExt	=> q_etDiagExt,
									q_sMsg		=> q_sMsg);

	IF q_etDiag <> GD.ET_Diag.Ok THEN
		RETURN;
	END_IF

THIS^.fbTreeWriter.NodeEnd(	q_etDiag	=> q_etDiag,
							q_etDiagExt	=> q_etDiagExt,
							q_sMsg		=> q_sMsg);

IF q_etDiag <> GD.ET_Diag.Ok THEN
	RETURN;
END_IF

(* ---- WriteInterfaceEnd.meth.st ---- *)
{attribute 'conditionalshow_all_locals'}
METHOD INTERNAL WriteInterfaceEnd : BOOL
VAR_INPUT
END_VAR
VAR_OUTPUT
	q_etDiag		: GD.ET_Diag;
	q_etDiagExt	: TPL.ET_DiagExt;
	q_sMsg			: STRING[80];
END_VAR

THIS^.fbTreeWriter.NodeEnd(	q_etDiag	=> q_etDiag,
							q_etDiagExt	=> q_etDiagExt,
							q_sMsg		=> q_sMsg);

(* ---- WriteInterfaceEndless.meth.st ---- *)
{attribute 'conditionalshow_all_locals'}
METHOD INTERNAL WriteInterfaceEndless : BOOL
VAR_INPUT
END_VAR
VAR_OUTPUT
	q_etDiag		: GD.ET_Diag;
	q_etDiagExt	: TPL.ET_DiagExt;
	q_sMsg			: STRING[80];
END_VAR

THIS^.fbTreeWriter.NodeStart(	i_sName		:= 'stEndless',
								q_etDiag	=> q_etDiag,
								q_etDiagExt	=> q_etDiagExt,
								q_sMsg		=> q_sMsg);

IF q_etDiag <> GD.ET_Diag.Ok THEN
	RETURN;
END_IF

	THIS^.fbTreeWriter.Parameter(	i_sName		:= 'i_lrVel',
									i_sValue	:= LREAL_TO_STRING(THIS^.pstInterface^.stEndless.i_lrVel),
									q_etDiag	=> q_etDiag,
									q_etDiagExt	=> q_etDiagExt,
									q_sMsg		=> q_sMsg);

	IF q_etDiag <> GD.ET_Diag.Ok THEN
		RETURN;
	END_IF

	THIS^.fbTreeWriter.Parameter(	i_sName		:= 'i_lrAcc',
									i_sValue	:= LREAL_TO_STRING(THIS^.pstInterface^.stEndless.i_lrAcc),
									q_etDiag	=> q_etDiag,
									q_etDiagExt	=> q_etDiagExt,
									q_sMsg		=> q_sMsg);

	IF q_etDiag <> GD.ET_Diag.Ok THEN
		RETURN;
	END_IF

	THIS^.fbTreeWriter.Parameter(	i_sName		:= 'i_lrDec',
									i_sValue	:= LREAL_TO_STRING(THIS^.pstInterface^.stEndless.i_lrDec),
									q_etDiag	=> q_etDiag,
									q_etDiagExt	=> q_etDiagExt,
									q_sMsg		=> q_sMsg);

	IF q_etDiag <> GD.ET_Diag.Ok THEN
		RETURN;
	END_IF

	THIS^.fbTreeWriter.Parameter(	i_sName		:= 'i_lrJerk',
									i_sValue	:= LREAL_TO_STRING(THIS^.pstInterface^.stEndless.i_lrJerk),
									q_etDiag	=> q_etDiag,
									q_etDiagExt	=> q_etDiagExt,
									q_sMsg		=> q_sMsg);

	IF q_etDiag <> GD.ET_Diag.Ok THEN
		RETURN;
	END_IF

	THIS^.fbTreeWriter.Parameter(	i_sName		:= 'i_lrPeriod',
									i_sValue	:= LREAL_TO_STRING(THIS^.pstInterface^.stEndless.i_lrPeriod),
									q_etDiag	=> q_etDiag,
									q_etDiagExt	=> q_etDiagExt,
									q_sMsg		=> q_sMsg);

	IF q_etDiag <> GD.ET_Diag.Ok THEN
		RETURN;
	END_IF

	THIS^.fbTreeWriter.Parameter(	i_sName		:= 'i_lrStopPosition',
									i_sValue	:= LREAL_TO_STRING(THIS^.pstInterface^.stEndless.i_lrStopPosition),
									q_etDiag	=> q_etDiag,
									q_etDiagExt	=> q_etDiagExt,
									q_sMsg		=> q_sMsg);

	IF q_etDiag <> GD.ET_Diag.Ok THEN
		RETURN;
	END_IF

	THIS^.fbTreeWriter.Parameter(	i_sName		:= 'q_xInVelocity',
									i_sValue	:= BOOL_TO_STRING(THIS^.pstInterface^.stEndless.q_xInVelocity),
									q_etDiag	=> q_etDiag,
									q_etDiagExt	=> q_etDiagExt,
									q_sMsg		=> q_sMsg);

	IF q_etDiag <> GD.ET_Diag.Ok THEN
		RETURN;
	END_IF

THIS^.fbTreeWriter.NodeEnd(	q_etDiag	=> q_etDiag,
							q_etDiagExt	=> q_etDiagExt,
							q_sMsg		=> q_sMsg);

IF q_etDiag <> GD.ET_Diag.Ok THEN
	RETURN;
END_IF

(* ---- WriteInterfaceHomeEnd.meth.st ---- *)
{attribute 'conditionalshow_all_locals'}
METHOD INTERNAL WriteInterfaceHomeEnd : BOOL
VAR_INPUT
END_VAR
VAR_OUTPUT
	q_etDiag		: GD.ET_Diag;
	q_etDiagExt	: TPL.ET_DiagExt;
	q_sMsg			: STRING[80];
END_VAR

THIS^.fbTreeWriter.NodeEnd(	q_etDiag	=> q_etDiag,
							q_etDiagExt	=> q_etDiagExt,
							q_sMsg		=> q_sMsg);

(* ---- WriteInterfaceHomeForce.meth.st ---- *)
{attribute 'conditionalshow_all_locals'}
METHOD INTERNAL WriteInterfaceHomeForce : BOOL
VAR_INPUT
END_VAR
VAR_OUTPUT
	q_etDiag		: GD.ET_Diag;
	q_etDiagExt	: TPL.ET_DiagExt;
	q_sMsg			: STRING[80];
END_VAR

THIS^.fbTreeWriter.NodeStart(	i_sName		:= 'stForce',
								q_etDiag	=> q_etDiag,
								q_etDiagExt	=> q_etDiagExt,
								q_sMsg		=> q_sMsg);

IF q_etDiag <> GD.ET_Diag.Ok THEN
	RETURN;
END_IF

	THIS^.fbTreeWriter.Parameter(	i_sName		:= 'i_lrHomePosition',
									i_sValue	:= LREAL_TO_STRING(THIS^.pstInterface^.stHome.stForce.i_lrHomePosition),
									q_etDiag	=> q_etDiag,
									q_etDiagExt	=> q_etDiagExt,
									q_sMsg		=> q_sMsg);

	IF q_etDiag <> GD.ET_Diag.Ok THEN
		RETURN;
	END_IF

	THIS^.fbTreeWriter.Parameter(	i_sName		:= 'i_lrVel',
									i_sValue	:= LREAL_TO_STRING(THIS^.pstInterface^.stHome.stForce.i_lrVel),
									q_etDiag	=> q_etDiag,
									q_etDiagExt	=> q_etDiagExt,
									q_sMsg		=> q_sMsg);

	IF q_etDiag <> GD.ET_Diag.Ok THEN
		RETURN;
	END_IF

	THIS^.fbTreeWriter.Parameter(	i_sName		:= 'i_lrAcc',
									i_sValue	:= LREAL_TO_STRING(THIS^.pstInterface^.stHome.stForce.i_lrAcc),
									q_etDiag	=> q_etDiag,
									q_etDiagExt	=> q_etDiagExt,
									q_sMsg		=> q_sMsg);

	IF q_etDiag <> GD.ET_Diag.Ok THEN
		RETURN;
	END_IF

	THIS^.fbTreeWriter.Parameter(	i_sName		:= 'i_lrDec',
									i_sValue	:= LREAL_TO_STRING(THIS^.pstInterface^.stHome.stForce.i_lrDec),
									q_etDiag	=> q_etDiag,
									q_etDiagExt	=> q_etDiagExt,
									q_sMsg		=> q_sMsg);

	IF q_etDiag <> GD.ET_Diag.Ok THEN
		RETURN;
	END_IF

	THIS^.fbTreeWriter.Parameter(	i_sName		:= 'i_lrJerk',
									i_sValue	:= LREAL_TO_STRING(THIS^.pstInterface^.stHome.stForce.i_lrJerk),
									q_etDiag	=> q_etDiag,
									q_etDiagExt	=> q_etDiagExt,
									q_sMsg		=> q_sMsg);

	IF q_etDiag <> GD.ET_Diag.Ok THEN
		RETURN;
	END_IF

	THIS^.fbTreeWriter.Parameter(	i_sName		:= 'i_lrOffset',
									i_sValue	:= LREAL_TO_STRING(THIS^.pstInterface^.stHome.stForce.i_lrOffset),
									q_etDiag	=> q_etDiag,
									q_etDiagExt	=> q_etDiagExt,
									q_sMsg		=> q_sMsg);

	IF q_etDiag <> GD.ET_Diag.Ok THEN
		RETURN;
	END_IF

	THIS^.fbTreeWriter.Parameter(	i_sName		:= 'i_lrMaxTravel',
									i_sValue	:= LREAL_TO_STRING(THIS^.pstInterface^.stHome.stForce.i_lrMaxTravel),
									q_etDiag	=> q_etDiag,
									q_etDiagExt	=> q_etDiagExt,
									q_sMsg		=> q_sMsg);

	IF q_etDiag <> GD.ET_Diag.Ok THEN
		RETURN;
	END_IF

	THIS^.fbTreeWriter.Parameter(	i_sName		:= 'i_lrMaxForce',
									i_sValue	:= LREAL_TO_STRING(THIS^.pstInterface^.stHome.stForce.i_lrMaxForce),
									q_etDiag	=> q_etDiag,
									q_etDiagExt	=> q_etDiagExt,
									q_sMsg		=> q_sMsg);

	IF q_etDiag <> GD.ET_Diag.Ok THEN
		RETURN;
	END_IF

	THIS^.fbTreeWriter.Parameter(	i_sName		:= 'i_diForceTime',
									i_sValue	:= DINT_TO_STRING(THIS^.pstInterface^.stHome.stForce.i_diForceTime),
									q_etDiag	=> q_etDiag,
									q_etDiagExt	=> q_etDiagExt,
									q_sMsg		=> q_sMsg);

	IF q_etDiag <> GD.ET_Diag.Ok THEN
		RETURN;
	END_IF

THIS^.fbTreeWriter.NodeEnd(	q_etDiag	=> q_etDiag,
							q_etDiagExt	=> q_etDiagExt,
							q_sMsg		=> q_sMsg);

IF q_etDiag <> GD.ET_Diag.Ok THEN
	RETURN;
END_IF

(* ---- WriteInterfaceHomeLimitSwitch.meth.st ---- *)
{attribute 'conditionalshow_all_locals'}
METHOD INTERNAL WriteInterfaceHomeLimitSwitch : BOOL
VAR_INPUT
END_VAR
VAR_OUTPUT
	q_etDiag		: GD.ET_Diag;
	q_etDiagExt	: TPL.ET_DiagExt;
	q_sMsg			: STRING[80];
END_VAR

THIS^.fbTreeWriter.NodeStart(	i_sName		:= 'stLimitSwitch',
								q_etDiag	=> q_etDiag,
								q_etDiagExt	=> q_etDiagExt,
								q_sMsg		=> q_sMsg);

IF q_etDiag <> GD.ET_Diag.Ok THEN
	RETURN;
END_IF

	THIS^.fbTreeWriter.Parameter(	i_sName		:= 'i_lrHomePosition',
									i_sValue	:= LREAL_TO_STRING(THIS^.pstInterface^.stHome.stLimitSwitch.i_lrHomePosition),
									q_etDiag	=> q_etDiag,
									q_etDiagExt	=> q_etDiagExt,
									q_sMsg		=> q_sMsg);

	IF q_etDiag <> GD.ET_Diag.Ok THEN
		RETURN;
	END_IF

	THIS^.fbTreeWriter.Parameter(	i_sName		:= 'i_lrVel',
									i_sValue	:= LREAL_TO_STRING(THIS^.pstInterface^.stHome.stLimitSwitch.i_lrVel),
									q_etDiag	=> q_etDiag,
									q_etDiagExt	=> q_etDiagExt,
									q_sMsg		=> q_sMsg);

	IF q_etDiag <> GD.ET_Diag.Ok THEN
		RETURN;
	END_IF

	THIS^.fbTreeWriter.Parameter(	i_sName		:= 'i_lrLowVel',
									i_sValue	:= LREAL_TO_STRING(THIS^.pstInterface^.stHome.stLimitSwitch.i_lrLowVel),
									q_etDiag	=> q_etDiag,
									q_etDiagExt	=> q_etDiagExt,
									q_sMsg		=> q_sMsg);

	IF q_etDiag <> GD.ET_Diag.Ok THEN
		RETURN;
	END_IF

	THIS^.fbTreeWriter.Parameter(	i_sName		:= 'i_lrAcc',
									i_sValue	:= LREAL_TO_STRING(THIS^.pstInterface^.stHome.stLimitSwitch.i_lrAcc),
									q_etDiag	=> q_etDiag,
									q_etDiagExt	=> q_etDiagExt,
									q_sMsg		=> q_sMsg);

	IF q_etDiag <> GD.ET_Diag.Ok THEN
		RETURN;
	END_IF

	THIS^.fbTreeWriter.Parameter(	i_sName		:= 'i_lrDec',
									i_sValue	:= LREAL_TO_STRING(THIS^.pstInterface^.stHome.stLimitSwitch.i_lrDec),
									q_etDiag	=> q_etDiag,
									q_etDiagExt	=> q_etDiagExt,
									q_sMsg		=> q_sMsg);

	IF q_etDiag <> GD.ET_Diag.Ok THEN
		RETURN;
	END_IF

	THIS^.fbTreeWriter.Parameter(	i_sName		:= 'i_lrJerk',
									i_sValue	:= LREAL_TO_STRING(THIS^.pstInterface^.stHome.stLimitSwitch.i_lrJerk),
									q_etDiag	=> q_etDiag,
									q_etDiagExt	=> q_etDiagExt,
									q_sMsg		=> q_sMsg);

	IF q_etDiag <> GD.ET_Diag.Ok THEN
		RETURN;
	END_IF

	THIS^.fbTreeWriter.Parameter(	i_sName		:= 'i_lrOffset',
									i_sValue	:= LREAL_TO_STRING(THIS^.pstInterface^.stHome.stLimitSwitch.i_lrOffset),
									q_etDiag	=> q_etDiag,
									q_etDiagExt	=> q_etDiagExt,
									q_sMsg		=> q_sMsg);

	IF q_etDiag <> GD.ET_Diag.Ok THEN
		RETURN;
	END_IF

	THIS^.fbTreeWriter.Parameter(	i_sName		:= 'i_lrMaxTravel',
									i_sValue	:= LREAL_TO_STRING(THIS^.pstInterface^.stHome.stLimitSwitch.i_lrMaxTravel),
									q_etDiag	=> q_etDiag,
									q_etDiagExt	=> q_etDiagExt,
									q_sMsg		=> q_sMsg);

	IF q_etDiag <> GD.ET_Diag.Ok THEN
		RETURN;
	END_IF

THIS^.fbTreeWriter.NodeEnd(	q_etDiag	=> q_etDiag,
							q_etDiagExt	=> q_etDiagExt,
							q_sMsg		=> q_sMsg);

IF q_etDiag <> GD.ET_Diag.Ok THEN
	RETURN;
END_IF

(* ---- WriteInterfaceHomeMoveOnPos.meth.st ---- *)
{attribute 'conditionalshow_all_locals'}
METHOD INTERNAL WriteInterfaceHomeMoveOnPos : BOOL
VAR_INPUT
END_VAR
VAR_OUTPUT
	q_etDiag		: GD.ET_Diag;
	q_etDiagExt	: TPL.ET_DiagExt;
	q_sMsg			: STRING[80];
END_VAR

THIS^.fbTreeWriter.NodeStart(	i_sName		:= 'stMoveOnPos',
								q_etDiag	=> q_etDiag,
								q_etDiagExt	=> q_etDiagExt,
								q_sMsg		=> q_sMsg);

IF q_etDiag <> GD.ET_Diag.Ok THEN
	RETURN;
END_IF

	THIS^.fbTreeWriter.Parameter(	i_sName		:= 'i_lrTarget',
									i_sValue	:= LREAL_TO_STRING(THIS^.pstInterface^.stHome.stMoveOnPos.i_lrTarget),
									q_etDiag	=> q_etDiag,
									q_etDiagExt	=> q_etDiagExt,
									q_sMsg		=> q_sMsg);

	IF q_etDiag <> GD.ET_Diag.Ok THEN
		RETURN;
	END_IF

	THIS^.fbTreeWriter.Parameter(	i_sName		:= 'i_lrVel',
									i_sValue	:= LREAL_TO_STRING(THIS^.pstInterface^.stHome.stMoveOnPos.i_lrVel),
									q_etDiag	=> q_etDiag,
									q_etDiagExt	=> q_etDiagExt,
									q_sMsg		=> q_sMsg);

	IF q_etDiag <> GD.ET_Diag.Ok THEN
		RETURN;
	END_IF

	THIS^.fbTreeWriter.Parameter(	i_sName		:= 'i_lrAcc',
									i_sValue	:= LREAL_TO_STRING(THIS^.pstInterface^.stHome.stMoveOnPos.i_lrAcc),
									q_etDiag	=> q_etDiag,
									q_etDiagExt	=> q_etDiagExt,
									q_sMsg		=> q_sMsg);

	IF q_etDiag <> GD.ET_Diag.Ok THEN
		RETURN;
	END_IF

	THIS^.fbTreeWriter.Parameter(	i_sName		:= 'i_lrDec',
									i_sValue	:= LREAL_TO_STRING(THIS^.pstInterface^.stHome.stMoveOnPos.i_lrDec),
									q_etDiag	=> q_etDiag,
									q_etDiagExt	=> q_etDiagExt,
									q_sMsg		=> q_sMsg);

	IF q_etDiag <> GD.ET_Diag.Ok THEN
		RETURN;
	END_IF

	THIS^.fbTreeWriter.Parameter(	i_sName		:= 'i_lrJerk',
									i_sValue	:= LREAL_TO_STRING(THIS^.pstInterface^.stHome.stMoveOnPos.i_lrJerk),
									q_etDiag	=> q_etDiag,
									q_etDiagExt	=> q_etDiagExt,
									q_sMsg		=> q_sMsg);

	IF q_etDiag <> GD.ET_Diag.Ok THEN
		RETURN;
	END_IF

	THIS^.fbTreeWriter.Parameter(	i_sName		:= 'i_xRotativeSystem',
									i_sValue	:= BOOL_TO_STRING(THIS^.pstInterface^.stHome.stMoveOnPos.i_xRotativeSystem),
									q_etDiag	=> q_etDiag,
									q_etDiagExt	=> q_etDiagExt,
									q_sMsg		=> q_sMsg);

	IF q_etDiag <> GD.ET_Diag.Ok THEN
		RETURN;
	END_IF

	THIS^.fbTreeWriter.Parameter(	i_sName		:= 'i_lrPeriod',
									i_sValue	:= LREAL_TO_STRING(THIS^.pstInterface^.stHome.stMoveOnPos.i_lrPeriod),
									q_etDiag	=> q_etDiag,
									q_etDiagExt	=> q_etDiagExt,
									q_sMsg		=> q_sMsg);

	IF q_etDiag <> GD.ET_Diag.Ok THEN
		RETURN;
	END_IF

THIS^.fbTreeWriter.NodeEnd(	q_etDiag	=> q_etDiag,
							q_etDiagExt	=> q_etDiagExt,
							q_sMsg		=> q_sMsg);

IF q_etDiag <> GD.ET_Diag.Ok THEN
	RETURN;
END_IF

(* ---- WriteInterfaceHomeParam.meth.st ---- *)
{attribute 'conditionalshow_all_locals'}
METHOD INTERNAL WriteInterfaceHomeParam : BOOL
VAR_INPUT
END_VAR
VAR_OUTPUT
	q_etDiag		: GD.ET_Diag;
	q_etDiagExt	: TPL.ET_DiagExt;
	q_sMsg			: STRING[80];
END_VAR

THIS^.fbTreeWriter.Parameter(	i_sName		:= 'i_xEnableInitAbsReadPos',
								i_sValue	:= BOOL_TO_STRING(THIS^.pstInterface^.stHome.i_xEnableInitAbsReadPos),
								q_etDiag	=> q_etDiag,
								q_etDiagExt	=> q_etDiagExt,
								q_sMsg		=> q_sMsg);

IF q_etDiag <> GD.ET_Diag.Ok THEN
	RETURN;
END_IF

THIS^.fbTreeWriter.Parameter(	i_sName		:= 'i_xResetHomeOk',
								i_sValue	:= BOOL_TO_STRING(THIS^.pstInterface^.stHome.i_xResetHomeOk),
								q_etDiag	=> q_etDiag,
								q_etDiagExt	=> q_etDiagExt,
								q_sMsg		=> q_sMsg);

IF q_etDiag <> GD.ET_Diag.Ok THEN
	RETURN;
END_IF

THIS^.fbTreeWriter.Parameter(	i_sName		:= 'i_etMode',
								i_sValue	:= AXM_FC_EtHomeModeToString(THIS^.pstInterface^.stHome.i_etMode),
								q_etDiag	=> q_etDiag,
								q_etDiagExt	=> q_etDiagExt,
								q_sMsg		=> q_sMsg);

IF q_etDiag <> GD.ET_Diag.Ok THEN
	RETURN;
END_IF

(* ---- WriteInterfaceHomeSensor.meth.st ---- *)
{attribute 'conditionalshow_all_locals'}
METHOD INTERNAL WriteInterfaceHomeSensor : BOOL
VAR_INPUT
END_VAR
VAR_OUTPUT
	q_etDiag		: GD.ET_Diag;
	q_etDiagExt	: TPL.ET_DiagExt;
	q_sMsg			: STRING[80];
END_VAR

THIS^.fbTreeWriter.NodeStart(	i_sName		:= 'stSensor',
								q_etDiag	=> q_etDiag,
								q_etDiagExt	=> q_etDiagExt,
								q_sMsg		=> q_sMsg);

IF q_etDiag <> GD.ET_Diag.Ok THEN
	RETURN;
END_IF

	THIS^.fbTreeWriter.Parameter(	i_sName		:= 'i_lrHomePosition',
									i_sValue	:= LREAL_TO_STRING(THIS^.pstInterface^.stHome.stSensor.i_lrHomePosition),
									q_etDiag	=> q_etDiag,
									q_etDiagExt	=> q_etDiagExt,
									q_sMsg		=> q_sMsg);

	IF q_etDiag <> GD.ET_Diag.Ok THEN
		RETURN;
	END_IF

	THIS^.fbTreeWriter.Parameter(	i_sName		:= 'i_lrVel',
									i_sValue	:= LREAL_TO_STRING(THIS^.pstInterface^.stHome.stSensor.i_lrVel),
									q_etDiag	=> q_etDiag,
									q_etDiagExt	=> q_etDiagExt,
									q_sMsg		=> q_sMsg);

	IF q_etDiag <> GD.ET_Diag.Ok THEN
		RETURN;
	END_IF

	THIS^.fbTreeWriter.Parameter(	i_sName		:= 'i_lrAcc',
									i_sValue	:= LREAL_TO_STRING(THIS^.pstInterface^.stHome.stSensor.i_lrAcc),
									q_etDiag	=> q_etDiag,
									q_etDiagExt	=> q_etDiagExt,
									q_sMsg		=> q_sMsg);

	IF q_etDiag <> GD.ET_Diag.Ok THEN
		RETURN;
	END_IF

	THIS^.fbTreeWriter.Parameter(	i_sName		:= 'i_lrDec',
									i_sValue	:= LREAL_TO_STRING(THIS^.pstInterface^.stHome.stSensor.i_lrDec),
									q_etDiag	=> q_etDiag,
									q_etDiagExt	=> q_etDiagExt,
									q_sMsg		=> q_sMsg);

	IF q_etDiag <> GD.ET_Diag.Ok THEN
		RETURN;
	END_IF

	THIS^.fbTreeWriter.Parameter(	i_sName		:= 'i_lrJerk',
									i_sValue	:= LREAL_TO_STRING(THIS^.pstInterface^.stHome.stSensor.i_lrJerk),
									q_etDiag	=> q_etDiag,
									q_etDiagExt	=> q_etDiagExt,
									q_sMsg		=> q_sMsg);

	IF q_etDiag <> GD.ET_Diag.Ok THEN
		RETURN;
	END_IF

	THIS^.fbTreeWriter.Parameter(	i_sName		:= 'i_lrOffset',
									i_sValue	:= LREAL_TO_STRING(THIS^.pstInterface^.stHome.stSensor.i_lrOffset),
									q_etDiag	=> q_etDiag,
									q_etDiagExt	=> q_etDiagExt,
									q_sMsg		=> q_sMsg);

	IF q_etDiag <> GD.ET_Diag.Ok THEN
		RETURN;
	END_IF

	THIS^.fbTreeWriter.Parameter(	i_sName		:= 'i_lrMaxTravel',
									i_sValue	:= LREAL_TO_STRING(THIS^.pstInterface^.stHome.stSensor.i_lrMaxTravel),
									q_etDiag	=> q_etDiag,
									q_etDiagExt	=> q_etDiagExt,
									q_sMsg		=> q_sMsg);

	IF q_etDiag <> GD.ET_Diag.Ok THEN
		RETURN;
	END_IF

	THIS^.fbTreeWriter.Parameter(	i_sName		:= 'i_xRotativeSystem',
									i_sValue	:= BOOL_TO_STRING(THIS^.pstInterface^.stHome.stSensor.i_xRotativeSystem),
									q_etDiag	=> q_etDiag,
									q_etDiagExt	=> q_etDiagExt,
									q_sMsg		=> q_sMsg);

	IF q_etDiag <> GD.ET_Diag.Ok THEN
		RETURN;
	END_IF

	THIS^.fbTreeWriter.Parameter(	i_sName		:= 'i_xSensor',
									i_sValue	:= BOOL_TO_STRING(THIS^.pstInterface^.stHome.stSensor.i_xSensor),
									q_etDiag	=> q_etDiag,
									q_etDiagExt	=> q_etDiagExt,
									q_sMsg		=> q_sMsg);

	IF q_etDiag <> GD.ET_Diag.Ok THEN
		RETURN;
	END_IF

THIS^.fbTreeWriter.NodeEnd(	q_etDiag	=> q_etDiag,
							q_etDiagExt	=> q_etDiagExt,
							q_sMsg		=> q_sMsg);

IF q_etDiag <> GD.ET_Diag.Ok THEN
	RETURN;
END_IF

(* ---- WriteInterfaceHomeSetPos.meth.st ---- *)
{attribute 'conditionalshow_all_locals'}
METHOD INTERNAL WriteInterfaceHomeSetPos : BOOL
VAR_INPUT
END_VAR
VAR_OUTPUT
	q_etDiag		: GD.ET_Diag;
	q_etDiagExt	: TPL.ET_DiagExt;
	q_sMsg			: STRING[80];
END_VAR

THIS^.fbTreeWriter.NodeStart(	i_sName		:= 'stSetPos',
								q_etDiag	=> q_etDiag,
								q_etDiagExt	=> q_etDiagExt,
								q_sMsg		=> q_sMsg);

IF q_etDiag <> GD.ET_Diag.Ok THEN
	RETURN;
END_IF

	THIS^.fbTreeWriter.Parameter(	i_sName		:= 'i_lrHomePosition',
									i_sValue	:= LREAL_TO_STRING(THIS^.pstInterface^.stHome.stSetPos.i_lrHomePosition),
									q_etDiag	=> q_etDiag,
									q_etDiagExt	=> q_etDiagExt,
									q_sMsg		=> q_sMsg);

	IF q_etDiag <> GD.ET_Diag.Ok THEN
		RETURN;
	END_IF

// 	THIS^.fbTreeWriter.Parameter(	i_sName		:= 'i_lrEncoderPosition',
// 									i_sValue	:= LREAL_TO_STRING(THIS^.pstInterface^.stHome.stSetPos.i_lrEncoderPosition),
// 									q_etDiag	=> q_etDiag,
// 									q_etDiagExt	=> q_etDiagExt,
// 									q_sMsg		=> q_sMsg);
//
// 	IF q_etDiag <> GD.ET_Diag.Ok THEN
// 		RETURN;
// 	END_IF
//
// 	THIS^.fbTreeWriter.Parameter(	i_sName		:= 'i_lrUserPeriod',
// 									i_sValue	:= LREAL_TO_STRING(THIS^.pstInterface^.stHome.stSetPos.i_lrUserPeriod),
// 									q_etDiag	=> q_etDiag,
// 									q_etDiagExt	=> q_etDiagExt,
// 									q_sMsg		=> q_sMsg);
//
// 	IF q_etDiag <> GD.ET_Diag.Ok THEN
// 		RETURN;
// 	END_IF
//
// 	THIS^.fbTreeWriter.Parameter(	i_sName		:= 'i_lrAbsEncOffset',
// 									i_sValue	:= LREAL_TO_STRING(THIS^.pstInterface^.stHome.stSetPos.i_lrAbsEncOffset),
// 									q_etDiag	=> q_etDiag,
// 									q_etDiagExt	=> q_etDiagExt,
// 									q_sMsg		=> q_sMsg);
//
// 	IF q_etDiag <> GD.ET_Diag.Ok THEN
// 		RETURN;
// 	END_IF
//
// 	THIS^.fbTreeWriter.Parameter(	i_sName		:= 'i_lrRestoreWindow',
// 									i_sValue	:= LREAL_TO_STRING(THIS^.pstInterface^.stHome.stSetPos.i_lrRestoreWindow),
// 									q_etDiag	=> q_etDiag,
// 									q_etDiagExt	=> q_etDiagExt,
// 									q_sMsg		=> q_sMsg);
//
// 	IF q_etDiag <> GD.ET_Diag.Ok THEN
// 		RETURN;
// 	END_IF
//
// 	IF (THIS^.pstInterface^.stHome.stSetPos.iq_pstRestorePosRetain <> 0) THEN
//
// 		THIS^.fbTreeWriter.NodeStart(	i_sName		:= 'iq_pstRestorePosRetain',
// 										q_etDiag	=> q_etDiag,
// 										q_etDiagExt	=> q_etDiagExt,
// 										q_sMsg		=> q_sMsg);
//
// 		IF q_etDiag <> GD.ET_Diag.Ok THEN
// 			RETURN;
// 		END_IF
//
// 			THIS^.fbTreeWriter.Parameter(	i_sName		:= 'lrEncPosition',
// 											i_sValue	:= LREAL_TO_STRING(THIS^.pstInterface^.stHome.stSetPos.iq_pstRestorePosRetain^.lrEncPosition),
// 											q_etDiag	=> q_etDiag,
// 											q_etDiagExt	=> q_etDiagExt,
// 											q_sMsg		=> q_sMsg);
//
// 			IF q_etDiag <> GD.ET_Diag.Ok THEN
// 				RETURN;
// 			END_IF
//
// 			THIS^.fbTreeWriter.Parameter(	i_sName		:= 'lrAxisPosition',
// 											i_sValue	:= LREAL_TO_STRING(THIS^.pstInterface^.stHome.stSetPos.iq_pstRestorePosRetain^.lrAxisPosition),
// 											q_etDiag	=> q_etDiag,
// 											q_etDiagExt	=> q_etDiagExt,
// 											q_sMsg		=> q_sMsg);
//
// 			IF q_etDiag <> GD.ET_Diag.Ok THEN
// 				RETURN;
// 			END_IF
//
// 			THIS^.fbTreeWriter.Parameter(	i_sName		:= 'lrCheckSum',
// 											i_sValue	:= LREAL_TO_STRING(THIS^.pstInterface^.stHome.stSetPos.iq_pstRestorePosRetain^.lrCheckSum),
// 											q_etDiag	=> q_etDiag,
// 											q_etDiagExt	=> q_etDiagExt,
// 											q_sMsg		=> q_sMsg);
//
// 			IF q_etDiag <> GD.ET_Diag.Ok THEN
// 				RETURN;
// 			END_IF
//
// 		THIS^.fbTreeWriter.NodeEnd(	q_etDiag	=> q_etDiag,
// 									q_etDiagExt	=> q_etDiagExt,
// 									q_sMsg		=> q_sMsg);
//
// 		IF q_etDiag <> GD.ET_Diag.Ok THEN
// 			RETURN;
// 		END_IF
//
// 	ELSE
// 		THIS^.fbTreeWriter.Parameter(	i_sName		:= 'iq_pstRestorePosRetain',
// 										i_sValue	:= 'not configured',
// 										q_etDiag	=> q_etDiag,
// 										q_etDiagExt	=> q_etDiagExt,
// 										q_sMsg		=> q_sMsg);
//
// 		IF q_etDiag <> GD.ET_Diag.Ok THEN
// 			RETURN;
// 		END_IF
// 	END_IF

THIS^.fbTreeWriter.NodeEnd(	q_etDiag	=> q_etDiag,
							q_etDiagExt	=> q_etDiagExt,
							q_sMsg		=> q_sMsg);

IF q_etDiag <> GD.ET_Diag.Ok THEN
	RETURN;
END_IF

(* ---- WriteInterfaceHomeStart.meth.st ---- *)
{attribute 'conditionalshow_all_locals'}
METHOD INTERNAL WriteInterfaceHomeStart : BOOL
VAR_INPUT
END_VAR
VAR_OUTPUT
	q_etDiag		: GD.ET_Diag;
	q_etDiagExt	: TPL.ET_DiagExt;
	q_sMsg			: STRING[80];
END_VAR

THIS^.fbTreeWriter.NodeStart(	i_sName		:= 'stHome',
								q_etDiag	=> q_etDiag,
								q_etDiagExt	=> q_etDiagExt,
								q_sMsg		=> q_sMsg);

(* ---- WriteInterfaceHomeTorque.meth.st ---- *)
{attribute 'conditionalshow_all_locals'}
METHOD INTERNAL WriteInterfaceHomeTorque : BOOL
VAR_INPUT
END_VAR
VAR_OUTPUT
	q_etDiag		: GD.ET_Diag;
	q_etDiagExt	: TPL.ET_DiagExt;
	q_sMsg			: STRING[80];
END_VAR

THIS^.fbTreeWriter.NodeStart(	i_sName		:= 'stTorque',
								q_etDiag	=> q_etDiag,
								q_etDiagExt	=> q_etDiagExt,
								q_sMsg		=> q_sMsg);

IF q_etDiag <> GD.ET_Diag.Ok THEN
	RETURN;
END_IF

	THIS^.fbTreeWriter.Parameter(	i_sName		:= 'i_lrHomePosition',
									i_sValue	:= LREAL_TO_STRING(THIS^.pstInterface^.stHome.stTorque.i_lrHomePosition),
									q_etDiag	=> q_etDiag,
									q_etDiagExt	=> q_etDiagExt,
									q_sMsg		=> q_sMsg);

	IF q_etDiag <> GD.ET_Diag.Ok THEN
		RETURN;
	END_IF

	THIS^.fbTreeWriter.Parameter(	i_sName		:= 'i_lrVel',
									i_sValue	:= LREAL_TO_STRING(THIS^.pstInterface^.stHome.stTorque.i_lrVel),
									q_etDiag	=> q_etDiag,
									q_etDiagExt	=> q_etDiagExt,
									q_sMsg		=> q_sMsg);

	IF q_etDiag <> GD.ET_Diag.Ok THEN
		RETURN;
	END_IF

	THIS^.fbTreeWriter.Parameter(	i_sName		:= 'i_lrAcc',
									i_sValue	:= LREAL_TO_STRING(THIS^.pstInterface^.stHome.stTorque.i_lrAcc),
									q_etDiag	=> q_etDiag,
									q_etDiagExt	=> q_etDiagExt,
									q_sMsg		=> q_sMsg);

	IF q_etDiag <> GD.ET_Diag.Ok THEN
		RETURN;
	END_IF

	THIS^.fbTreeWriter.Parameter(	i_sName		:= 'i_lrDec',
									i_sValue	:= LREAL_TO_STRING(THIS^.pstInterface^.stHome.stTorque.i_lrDec),
									q_etDiag	=> q_etDiag,
									q_etDiagExt	=> q_etDiagExt,
									q_sMsg		=> q_sMsg);

	IF q_etDiag <> GD.ET_Diag.Ok THEN
		RETURN;
	END_IF

	THIS^.fbTreeWriter.Parameter(	i_sName		:= 'i_lrJerk',
									i_sValue	:= LREAL_TO_STRING(THIS^.pstInterface^.stHome.stTorque.i_lrJerk),
									q_etDiag	=> q_etDiag,
									q_etDiagExt	=> q_etDiagExt,
									q_sMsg		=> q_sMsg);

	IF q_etDiag <> GD.ET_Diag.Ok THEN
		RETURN;
	END_IF

	THIS^.fbTreeWriter.Parameter(	i_sName		:= 'i_lrOffset',
									i_sValue	:= LREAL_TO_STRING(THIS^.pstInterface^.stHome.stTorque.i_lrOffset),
									q_etDiag	=> q_etDiag,
									q_etDiagExt	=> q_etDiagExt,
									q_sMsg		=> q_sMsg);

	IF q_etDiag <> GD.ET_Diag.Ok THEN
		RETURN;
	END_IF

	THIS^.fbTreeWriter.Parameter(	i_sName		:= 'i_lrMaxTravel',
									i_sValue	:= LREAL_TO_STRING(THIS^.pstInterface^.stHome.stTorque.i_lrMaxTravel),
									q_etDiag	=> q_etDiag,
									q_etDiagExt	=> q_etDiagExt,
									q_sMsg		=> q_sMsg);

	IF q_etDiag <> GD.ET_Diag.Ok THEN
		RETURN;
	END_IF

	THIS^.fbTreeWriter.Parameter(	i_sName		:= 'i_lrMaxTorque',
									i_sValue	:= LREAL_TO_STRING(THIS^.pstInterface^.stHome.stTorque.i_lrMaxTorque),
									q_etDiag	=> q_etDiag,
									q_etDiagExt	=> q_etDiagExt,
									q_sMsg		=> q_sMsg);

	IF q_etDiag <> GD.ET_Diag.Ok THEN
		RETURN;
	END_IF

	THIS^.fbTreeWriter.Parameter(	i_sName		:= 'i_diTorqueTime',
									i_sValue	:= DINT_TO_STRING(THIS^.pstInterface^.stHome.stTorque.i_diTorqueTime),
									q_etDiag	=> q_etDiag,
									q_etDiagExt	=> q_etDiagExt,
									q_sMsg		=> q_sMsg);

	IF q_etDiag <> GD.ET_Diag.Ok THEN
		RETURN;
	END_IF

THIS^.fbTreeWriter.NodeEnd(	q_etDiag	=> q_etDiag,
							q_etDiagExt	=> q_etDiagExt,
							q_sMsg		=> q_sMsg);

IF q_etDiag <> GD.ET_Diag.Ok THEN
	RETURN;
END_IF

(* ---- WriteInterfaceHomeTouchProbe.meth.st ---- *)
{attribute 'conditionalshow_all_locals'}
METHOD INTERNAL WriteInterfaceHomeTouchProbe : BOOL
VAR_INPUT
END_VAR
VAR_OUTPUT
	q_etDiag		: GD.ET_Diag;
	q_etDiagExt	: TPL.ET_DiagExt;
	q_sMsg			: STRING[80];
END_VAR

THIS^.fbTreeWriter.NodeStart(	i_sName		:= 'stTouchProbe',
								q_etDiag	=> q_etDiag,
								q_etDiagExt	=> q_etDiagExt,
								q_sMsg		=> q_sMsg);

IF q_etDiag <> GD.ET_Diag.Ok THEN
	RETURN;
END_IF

	THIS^.fbTreeWriter.Parameter(	i_sName		:= 'i_lrHomePosition',
									i_sValue	:= LREAL_TO_STRING(THIS^.pstInterface^.stHome.stTouchProbe.i_lrHomePosition),
									q_etDiag	=> q_etDiag,
									q_etDiagExt	=> q_etDiagExt,
									q_sMsg		=> q_sMsg);

	IF q_etDiag <> GD.ET_Diag.Ok THEN
		RETURN;
	END_IF

	THIS^.fbTreeWriter.Parameter(	i_sName		:= 'i_lrVel',
									i_sValue	:= LREAL_TO_STRING(THIS^.pstInterface^.stHome.stTouchProbe.i_lrVel),
									q_etDiag	=> q_etDiag,
									q_etDiagExt	=> q_etDiagExt,
									q_sMsg		=> q_sMsg);

	IF q_etDiag <> GD.ET_Diag.Ok THEN
		RETURN;
	END_IF

	THIS^.fbTreeWriter.Parameter(	i_sName		:= 'i_lrAcc',
									i_sValue	:= LREAL_TO_STRING(THIS^.pstInterface^.stHome.stTouchProbe.i_lrAcc),
									q_etDiag	=> q_etDiag,
									q_etDiagExt	=> q_etDiagExt,
									q_sMsg		=> q_sMsg);

	IF q_etDiag <> GD.ET_Diag.Ok THEN
		RETURN;
	END_IF

	THIS^.fbTreeWriter.Parameter(	i_sName		:= 'i_lrDec',
									i_sValue	:= LREAL_TO_STRING(THIS^.pstInterface^.stHome.stTouchProbe.i_lrDec),
									q_etDiag	=> q_etDiag,
									q_etDiagExt	=> q_etDiagExt,
									q_sMsg		=> q_sMsg);

	IF q_etDiag <> GD.ET_Diag.Ok THEN
		RETURN;
	END_IF

	THIS^.fbTreeWriter.Parameter(	i_sName		:= 'i_lrJerk',
									i_sValue	:= LREAL_TO_STRING(THIS^.pstInterface^.stHome.stTouchProbe.i_lrJerk),
									q_etDiag	=> q_etDiag,
									q_etDiagExt	=> q_etDiagExt,
									q_sMsg		=> q_sMsg);

	IF q_etDiag <> GD.ET_Diag.Ok THEN
		RETURN;
	END_IF

	THIS^.fbTreeWriter.Parameter(	i_sName		:= 'i_lrOffset',
									i_sValue	:= LREAL_TO_STRING(THIS^.pstInterface^.stHome.stTouchProbe.i_lrOffset),
									q_etDiag	=> q_etDiag,
									q_etDiagExt	=> q_etDiagExt,
									q_sMsg		=> q_sMsg);

	IF q_etDiag <> GD.ET_Diag.Ok THEN
		RETURN;
	END_IF

	THIS^.fbTreeWriter.Parameter(	i_sName		:= 'i_lrMaxTravel',
									i_sValue	:= LREAL_TO_STRING(THIS^.pstInterface^.stHome.stTouchProbe.i_lrMaxTravel),
									q_etDiag	=> q_etDiag,
									q_etDiagExt	=> q_etDiagExt,
									q_sMsg		=> q_sMsg);

	IF q_etDiag <> GD.ET_Diag.Ok THEN
		RETURN;
	END_IF

	THIS^.fbTreeWriter.Parameter(	i_sName		:= 'i_xRotativeSystem',
									i_sValue	:= BOOL_TO_STRING(THIS^.pstInterface^.stHome.stTouchProbe.i_xRotativeSystem),
									q_etDiag	=> q_etDiag,
									q_etDiagExt	=> q_etDiagExt,
									q_sMsg		=> q_sMsg);

	IF q_etDiag <> GD.ET_Diag.Ok THEN
		RETURN;
	END_IF

// 	(* get drive name for variables i_ifDrive *)
// 	IF (THIS^.pstInterface^.stHome.stTouchProbe.i_ifTouchProbe <> 0) THEN
// 		THIS^.sTmp := THIS^.pstInterface^.stHome.stTouchProbe.i_ifTouchProbe.Name;
// 	ELSE
// 		THIS^.sTmp := 'not configured';
// 	END_IF
//
// 	THIS^.fbTreeWriter.Parameter(	i_sName		:= 'i_ifTouchProbe',
// 									i_sValue	:= THIS^.sTmp,
// 									q_etDiag	=> q_etDiag,
// 									q_etDiagExt	=> q_etDiagExt,
// 									q_sMsg		=> q_sMsg);
//
// 	IF q_etDiag <> GD.ET_Diag.Ok THEN
// 		RETURN;
// 	END_IF

THIS^.fbTreeWriter.NodeEnd(	q_etDiag	=> q_etDiag,
							q_etDiagExt	=> q_etDiagExt,
							q_sMsg		=> q_sMsg);

IF q_etDiag <> GD.ET_Diag.Ok THEN
	RETURN;
END_IF

(* ---- WriteInterfaceHomeWritePos.meth.st ---- *)
{attribute 'conditionalshow_all_locals'}
METHOD INTERNAL WriteInterfaceHomeWritePos : BOOL
VAR_INPUT
END_VAR
VAR_OUTPUT
	q_etDiag		: GD.ET_Diag;
	q_etDiagExt	: TPL.ET_DiagExt;
	q_sMsg			: STRING[80];
END_VAR

THIS^.fbTreeWriter.NodeStart(	i_sName		:= 'stWritePos',
								q_etDiag	=> q_etDiag,
								q_etDiagExt	=> q_etDiagExt,
								q_sMsg		=> q_sMsg);

IF q_etDiag <> GD.ET_Diag.Ok THEN
	RETURN;
END_IF

	THIS^.fbTreeWriter.Parameter(	i_sName		:= 'i_lrHomePosition',
									i_sValue	:= LREAL_TO_STRING(THIS^.pstInterface^.stHome.stWritePos.i_lrHomePosition),
									q_etDiag	=> q_etDiag,
									q_etDiagExt	=> q_etDiagExt,
									q_sMsg		=> q_sMsg);

	IF q_etDiag <> GD.ET_Diag.Ok THEN
		RETURN;
	END_IF

	THIS^.fbTreeWriter.Parameter(	i_sName		:= 'i_lrUserPeriod',
									i_sValue	:= LREAL_TO_STRING(THIS^.pstInterface^.stHome.stWritePos.i_lrUserPeriod),
									q_etDiag	=> q_etDiag,
									q_etDiagExt	=> q_etDiagExt,
									q_sMsg		=> q_sMsg);

	IF q_etDiag <> GD.ET_Diag.Ok THEN
		RETURN;
	END_IF

	THIS^.fbTreeWriter.Parameter(	i_sName		:= 'i_lrAbsEncOffset',
									i_sValue	:= LREAL_TO_STRING(THIS^.pstInterface^.stHome.stWritePos.i_lrAbsEncOffset),
									q_etDiag	=> q_etDiag,
									q_etDiagExt	=> q_etDiagExt,
									q_sMsg		=> q_sMsg);

	IF q_etDiag <> GD.ET_Diag.Ok THEN
		RETURN;
	END_IF

THIS^.fbTreeWriter.NodeEnd(	q_etDiag	=> q_etDiag,
							q_etDiagExt	=> q_etDiagExt,
							q_sMsg		=> q_sMsg);

IF q_etDiag <> GD.ET_Diag.Ok THEN
	RETURN;
END_IF

(* ---- WriteInterfaceMain.meth.st ---- *)
{attribute 'conditionalshow_all_locals'}
METHOD INTERNAL WriteInterfaceMain : BOOL
VAR_INPUT
END_VAR
VAR_OUTPUT
	q_etDiag		: GD.ET_Diag;
	q_etDiagExt	: TPL.ET_DiagExt;
	q_sMsg			: STRING[80];
END_VAR

THIS^.fbTreeWriter.NodeStart(	i_sName		:= 'stMain',
								q_etDiag	=> q_etDiag,
								q_etDiagExt	=> q_etDiagExt,
								q_sMsg		=> q_sMsg);

IF q_etDiag <> GD.ET_Diag.Ok THEN
	RETURN;
END_IF

// 	(* get drive name for variables i_ifDrive *)
// 	IF (THIS^.pstInterface^.stMain.i_ifDrive <> 0) THEN
// 		THIS^.sTmp := THIS^.pstInterface^.stMain.i_ifDrive.Name;
// 	ELSE
// 		THIS^.sTmp := 'not configured';
// 	END_IF
//
// 	THIS^.fbTreeWriter.Parameter(	i_sName		:= 'i_ifDrive',
// 									i_sValue	:= THIS^.sTmp,
// 									q_etDiag	=> q_etDiag,
// 									q_etDiagExt	=> q_etDiagExt,
// 									q_sMsg		=> q_sMsg);
//
// 	IF q_etDiag <> GD.ET_Diag.Ok THEN
// 		RETURN;
// 	END_IF

// 	(* get master name for variables i_ifMaster *)
// 	IF (THIS^.pstInterface^.stMain.i_ifMaster <> 0) THEN
// 		THIS^.sTmp := THIS^.pstInterface^.stMain.i_ifMaster.Name;
// 	ELSE
// 		THIS^.sTmp := 'not configured';
// 	END_IF
//
// 	THIS^.fbTreeWriter.Parameter(	i_sName		:= 'i_ifMaster',
// 									i_sValue	:= THIS^.sTmp,
// 									q_etDiag	=> q_etDiag,
// 									q_etDiagExt	=> q_etDiagExt,
// 									q_sMsg		=> q_sMsg);
//
// 	IF q_etDiag <> GD.ET_Diag.Ok THEN
// 		RETURN;
// 	END_IF

	THIS^.fbTreeWriter.Parameter(	i_sName		:= 'i_timMasterStop',
									i_sValue	:= TIME_TO_STRING(THIS^.pstInterface^.stMain.i_timMasterStop),
									q_etDiag	=> q_etDiag,
									q_etDiagExt	=> q_etDiagExt,
									q_sMsg		=> q_sMsg);

	IF q_etDiag <> GD.ET_Diag.Ok THEN
		RETURN;
	END_IF

	THIS^.fbTreeWriter.Parameter(	i_sName		:= 'i_xHwLimitPos',
									i_sValue	:= BOOL_TO_STRING(THIS^.pstInterface^.stMain.i_xHwLimitPos),
									q_etDiag	=> q_etDiag,
									q_etDiagExt	=> q_etDiagExt,
									q_sMsg		=> q_sMsg);

	IF q_etDiag <> GD.ET_Diag.Ok THEN
		RETURN;
	END_IF

	THIS^.fbTreeWriter.Parameter(	i_sName		:= 'i_xHwLimitNeg',
									i_sValue	:= BOOL_TO_STRING(THIS^.pstInterface^.stMain.i_xHwLimitNeg),
									q_etDiag	=> q_etDiag,
									q_etDiagExt	=> q_etDiagExt,
									q_sMsg		=> q_sMsg);

	IF q_etDiag <> GD.ET_Diag.Ok THEN
		RETURN;
	END_IF

	THIS^.fbTreeWriter.Parameter(	i_sName		:= 'i_xStart',
									i_sValue	:= BOOL_TO_STRING(THIS^.pstInterface^.stMain.i_xStart),
									q_etDiag	=> q_etDiag,
									q_etDiagExt	=> q_etDiagExt,
									q_sMsg		=> q_sMsg);

	IF q_etDiag <> GD.ET_Diag.Ok THEN
		RETURN;
	END_IF

	THIS^.fbTreeWriter.Parameter(	i_sName		:= 'i_lrMotionActiveVelLimit',
									i_sValue	:= LREAL_TO_STRING(THIS^.pstInterface^.stMain.i_lrMotionActiveVelLimit),
									q_etDiag	=> q_etDiag,
									q_etDiagExt	=> q_etDiagExt,
									q_sMsg		=> q_sMsg);

	IF q_etDiag <> GD.ET_Diag.Ok THEN
		RETURN;
	END_IF

	THIS^.fbTreeWriter.Parameter(	i_sName		:= 'i_etMotionActiveVelType',
									i_sValue	:= AXM_FC_EtMotionActiveVelTypeToString(THIS^.pstInterface^.stMain.i_etMotionActiveVelType),
									q_etDiag	=> q_etDiag,
									q_etDiagExt	=> q_etDiagExt,
									q_sMsg		=> q_sMsg);

	IF q_etDiag <> GD.ET_Diag.Ok THEN
		RETURN;
	END_IF

// 	(* get lenc name for variables iq_lencEncoder *)
// 	stLogicalAddress := THIS^.pstInterface^.stMain.iq_lencEncoder.stLogicalAddress;
// 	IF (stLogicalAddress.udiInstance <> 0) THEN
// 		THIS^.sTmp := THIS^.pstInterface^.stMain.iq_lencEncoder.Name;
// 	ELSE
// 		THIS^.sTmp := 'not configured';
// 	END_IF
//
// 	THIS^.fbTreeWriter.Parameter(	i_sName		:= 'iq_lencEncoder',
// 									i_sValue	:= THIS^.sTmp,
// 									q_etDiag	=> q_etDiag,
// 									q_etDiagExt	=> q_etDiagExt,
// 									q_sMsg		=> q_sMsg);
//
// 	IF q_etDiag <> GD.ET_Diag.Ok THEN
// 		RETURN;
// 	END_IF

	THIS^.fbTreeWriter.NodeStart(	i_sName		:= 'stReducedVelocity',
									q_etDiag	=> q_etDiag,
									q_etDiagExt	=> q_etDiagExt,
									q_sMsg		=> q_sMsg);

	IF q_etDiag <> GD.ET_Diag.Ok THEN
		RETURN;
	END_IF

		THIS^.fbTreeWriter.Parameter(	i_sName		:= 'i_xEnableReducedVelocity',
										i_sValue	:= BOOL_TO_STRING(THIS^.pstInterface^.stMain.stReducedVelocity.i_xEnableReducedVelocity),
										q_etDiag	=> q_etDiag,
										q_etDiagExt	=> q_etDiagExt,
										q_sMsg		=> q_sMsg);

		IF q_etDiag <> GD.ET_Diag.Ok THEN
			RETURN;
		END_IF

		THIS^.fbTreeWriter.Parameter(	i_sName		:= 'i_lrMaxReducedVelocity',
										i_sValue	:= LREAL_TO_STRING(THIS^.pstInterface^.stMain.stReducedVelocity.i_lrMaxReducedVelocity),
										q_etDiag	=> q_etDiag,
										q_etDiagExt	=> q_etDiagExt,
										q_sMsg		=> q_sMsg);

		IF q_etDiag <> GD.ET_Diag.Ok THEN
			RETURN;
		END_IF

		THIS^.fbTreeWriter.Parameter(	i_sName		:= 'i_xOnlyLimitCheck',
										i_sValue	:= BOOL_TO_STRING(THIS^.pstInterface^.stMain.stReducedVelocity.i_xOnlyLimitCheck),
										q_etDiag	=> q_etDiag,
										q_etDiagExt	=> q_etDiagExt,
										q_sMsg		=> q_sMsg);

		IF q_etDiag <> GD.ET_Diag.Ok THEN
			RETURN;
		END_IF

		THIS^.fbTreeWriter.Parameter(	i_sName		:= 'i_lrReducedVelocityCheckFactor',
										i_sValue	:= LREAL_TO_STRING(THIS^.pstInterface^.stMain.stReducedVelocity.i_lrReducedVelocityCheckFactor),
										q_etDiag	=> q_etDiag,
										q_etDiagExt	=> q_etDiagExt,
										q_sMsg		=> q_sMsg);

		IF q_etDiag <> GD.ET_Diag.Ok THEN
			RETURN;
		END_IF

	THIS^.fbTreeWriter.NodeEnd(	q_etDiag	=> q_etDiag,
								q_etDiagExt	=> q_etDiagExt,
								q_sMsg		=> q_sMsg);

	IF q_etDiag <> GD.ET_Diag.Ok THEN
		RETURN;
	END_IF

	THIS^.fbTreeWriter.Parameter(	i_sName		:= 'q_xDriveActive',
									i_sValue	:= BOOL_TO_STRING(THIS^.pstInterface^.stMain.q_xDriveActive),
									q_etDiag	=> q_etDiag,
									q_etDiagExt	=> q_etDiagExt,
									q_sMsg		=> q_sMsg);

	IF q_etDiag <> GD.ET_Diag.Ok THEN
		RETURN;
	END_IF

	THIS^.fbTreeWriter.Parameter(	i_sName		:= 'q_etOpMode',
									i_sValue	:= AXM_FC_EtOpModeToString(THIS^.pstInterface^.stMain.q_etOpMode),
									q_etDiag	=> q_etDiag,
									q_etDiagExt	=> q_etDiagExt,
									q_sMsg		=> q_sMsg);

	IF q_etDiag <> GD.ET_Diag.Ok THEN
		RETURN;
	END_IF

	THIS^.fbTreeWriter.Parameter(	i_sName		:= 'q_etState',
									i_sValue	:= AXM_FC_EtStateToString(THIS^.pstInterface^.stMain.q_etState),
									q_etDiag	=> q_etDiag,
									q_etDiagExt	=> q_etDiagExt,
									q_sMsg		=> q_sMsg);

	IF q_etDiag <> GD.ET_Diag.Ok THEN
		RETURN;
	END_IF

	THIS^.fbTreeWriter.Parameter(	i_sName		:= 'q_xHomeOk',
									i_sValue	:= BOOL_TO_STRING(THIS^.pstInterface^.stMain.q_xHomeOk),
									q_etDiag	=> q_etDiag,
									q_etDiagExt	=> q_etDiagExt,
									q_sMsg		=> q_sMsg);

	IF q_etDiag <> GD.ET_Diag.Ok THEN
		RETURN;
	END_IF

	THIS^.fbTreeWriter.Parameter(	i_sName		:= 'q_xSynchron',
									i_sValue	:= BOOL_TO_STRING(THIS^.pstInterface^.stMain.q_xSynchron),
									q_etDiag	=> q_etDiag,
									q_etDiagExt	=> q_etDiagExt,
									q_sMsg		=> q_sMsg);

	IF q_etDiag <> GD.ET_Diag.Ok THEN
		RETURN;
	END_IF

	THIS^.fbTreeWriter.Parameter(	i_sName		:= 'q_lrPosition',
									i_sValue	:= LREAL_TO_STRING(THIS^.pstInterface^.stMain.q_lrPosition),
									q_etDiag	=> q_etDiag,
									q_etDiagExt	=> q_etDiagExt,
									q_sMsg		=> q_sMsg);

	IF q_etDiag <> GD.ET_Diag.Ok THEN
		RETURN;
	END_IF

	THIS^.fbTreeWriter.Parameter(	i_sName		:= 'q_lrPositionX',
									i_sValue	:= LREAL_TO_STRING(THIS^.pstInterface^.stMain.q_lrPositionX),
									q_etDiag	=> q_etDiag,
									q_etDiagExt	=> q_etDiagExt,
									q_sMsg		=> q_sMsg);

	IF q_etDiag <> GD.ET_Diag.Ok THEN
		RETURN;
	END_IF

// 	THIS^.fbTreeWriter.Parameter(	i_sName		:= 'q_sDriveName',
// 									i_sValue	:= THIS^.pstInterface^.stMain.q_sDriveName,
// 									q_etDiag	=> q_etDiag,
// 									q_etDiagExt	=> q_etDiagExt,
// 									q_sMsg		=> q_sMsg);
//
// 	IF q_etDiag <> GD.ET_Diag.Ok THEN
// 		RETURN;
// 	END_IF

	THIS^.fbTreeWriter.Parameter(	i_sName		:= 'q_xMotionActive',
									i_sValue	:= BOOL_TO_STRING(THIS^.pstInterface^.stMain.q_xMotionActive),
									q_etDiag	=> q_etDiag,
									q_etDiagExt	=> q_etDiagExt,
									q_sMsg		=> q_sMsg);

	IF q_etDiag <> GD.ET_Diag.Ok THEN
		RETURN;
	END_IF

THIS^.fbTreeWriter.NodeEnd(	q_etDiag	=> q_etDiag,
							q_etDiagExt	=> q_etDiagExt,
							q_sMsg		=> q_sMsg);

IF q_etDiag <> GD.ET_Diag.Ok THEN
	RETURN;
END_IF

(* ---- WriteInterfaceManual.meth.st ---- *)
{attribute 'conditionalshow_all_locals'}
METHOD INTERNAL WriteInterfaceManual : BOOL
VAR_INPUT
END_VAR
VAR_OUTPUT
	q_etDiag		: GD.ET_Diag;
	q_etDiagExt	: TPL.ET_DiagExt;
	q_sMsg			: STRING[80];
END_VAR

THIS^.fbTreeWriter.NodeStart(	i_sName		:= 'stManual',
								q_etDiag	=> q_etDiag,
								q_etDiagExt	=> q_etDiagExt,
								q_sMsg		=> q_sMsg);

IF q_etDiag <> GD.ET_Diag.Ok THEN
	RETURN;
END_IF

	THIS^.fbTreeWriter.Parameter(	i_sName		:= 'i_xJogForw',
									i_sValue	:= BOOL_TO_STRING(THIS^.pstInterface^.stManual.i_xJogForw),
									q_etDiag	=> q_etDiag,
									q_etDiagExt	=> q_etDiagExt,
									q_sMsg		=> q_sMsg);

	IF q_etDiag <> GD.ET_Diag.Ok THEN
		RETURN;
	END_IF

	THIS^.fbTreeWriter.Parameter(	i_sName		:= 'i_xJogBack',
									i_sValue	:= BOOL_TO_STRING(THIS^.pstInterface^.stManual.i_xJogBack),
									q_etDiag	=> q_etDiag,
									q_etDiagExt	=> q_etDiagExt,
									q_sMsg		=> q_sMsg);

	IF q_etDiag <> GD.ET_Diag.Ok THEN
		RETURN;
	END_IF

	THIS^.fbTreeWriter.Parameter(	i_sName		:= 'i_lrVel',
									i_sValue	:= LREAL_TO_STRING(THIS^.pstInterface^.stManual.i_lrVel),
									q_etDiag	=> q_etDiag,
									q_etDiagExt	=> q_etDiagExt,
									q_sMsg		=> q_sMsg);

	IF q_etDiag <> GD.ET_Diag.Ok THEN
		RETURN;
	END_IF

	THIS^.fbTreeWriter.Parameter(	i_sName		:= 'i_lrAcc',
									i_sValue	:= LREAL_TO_STRING(THIS^.pstInterface^.stManual.i_lrAcc),
									q_etDiag	=> q_etDiag,
									q_etDiagExt	=> q_etDiagExt,
									q_sMsg		=> q_sMsg);

	IF q_etDiag <> GD.ET_Diag.Ok THEN
		RETURN;
	END_IF

	THIS^.fbTreeWriter.Parameter(	i_sName		:= 'i_lrDec',
									i_sValue	:= LREAL_TO_STRING(THIS^.pstInterface^.stManual.i_lrDec),
									q_etDiag	=> q_etDiag,
									q_etDiagExt	=> q_etDiagExt,
									q_sMsg		=> q_sMsg);

	IF q_etDiag <> GD.ET_Diag.Ok THEN
		RETURN;
	END_IF

	THIS^.fbTreeWriter.Parameter(	i_sName		:= 'i_lrJerk',
									i_sValue	:= LREAL_TO_STRING(THIS^.pstInterface^.stManual.i_lrJerk),
									q_etDiag	=> q_etDiag,
									q_etDiagExt	=> q_etDiagExt,
									q_sMsg		=> q_sMsg);

	IF q_etDiag <> GD.ET_Diag.Ok THEN
		RETURN;
	END_IF

	THIS^.fbTreeWriter.Parameter(	i_sName		:= 'i_lrMaxDistance',
									i_sValue	:= LREAL_TO_STRING(THIS^.pstInterface^.stManual.i_lrMaxDistance),
									q_etDiag	=> q_etDiag,
									q_etDiagExt	=> q_etDiagExt,
									q_sMsg		=> q_sMsg);

	IF q_etDiag <> GD.ET_Diag.Ok THEN
		RETURN;
	END_IF

	THIS^.fbTreeWriter.Parameter(	i_sName		:= 'i_lrPeriod',
									i_sValue	:= LREAL_TO_STRING(THIS^.pstInterface^.stManual.i_lrPeriod),
									q_etDiag	=> q_etDiag,
									q_etDiagExt	=> q_etDiagExt,
									q_sMsg		=> q_sMsg);

	IF q_etDiag <> GD.ET_Diag.Ok THEN
		RETURN;
	END_IF

	THIS^.fbTreeWriter.Parameter(	i_sName		:= 'i_xEndless',
									i_sValue	:= BOOL_TO_STRING(THIS^.pstInterface^.stManual.i_xEndless),
									q_etDiag	=> q_etDiag,
									q_etDiagExt	=> q_etDiagExt,
									q_sMsg		=> q_sMsg);

	IF q_etDiag <> GD.ET_Diag.Ok THEN
		RETURN;
	END_IF

THIS^.fbTreeWriter.NodeEnd(	q_etDiag	=> q_etDiag,
							q_etDiagExt	=> q_etDiagExt,
							q_sMsg		=> q_sMsg);

IF q_etDiag <> GD.ET_Diag.Ok THEN
	RETURN;
END_IF

(* ---- WriteInterfaceMultiCamEnd.meth.st ---- *)
{attribute 'conditionalshow_all_locals'}
METHOD INTERNAL WriteInterfaceMultiCamEnd : BOOL
VAR_INPUT
END_VAR
VAR_OUTPUT
	q_etDiag		: GD.ET_Diag;
	q_etDiagExt	: TPL.ET_DiagExt;
	q_sMsg			: STRING[80];
END_VAR

THIS^.fbTreeWriter.NodeEnd(	q_etDiag	=> q_etDiag,
							q_etDiagExt	=> q_etDiagExt,
							q_sMsg		=> q_sMsg);

(* ---- WriteInterfaceMultiCamExt.meth.st ---- *)
{attribute 'conditionalshow_all_locals'}
METHOD INTERNAL WriteInterfaceMultiCamExt : BOOL
VAR_INPUT
END_VAR
VAR_OUTPUT
	q_etDiag		: GD.ET_Diag;
	q_etDiagExt	: TPL.ET_DiagExt;
	q_sMsg			: STRING[80];
END_VAR

THIS^.fbTreeWriter.NodeStart(	i_sName		:= 'iq_stExt',
								q_etDiag	=> q_etDiag,
								q_etDiagExt	=> q_etDiagExt,
								q_sMsg		=> q_sMsg);

IF q_etDiag <> GD.ET_Diag.Ok THEN
	RETURN;
END_IF

	THIS^.fbTreeWriter.Parameter(	i_sName		:= 'xNoModuloMasterAtStart',
									i_sValue	:= BOOL_TO_STRING(THIS^.pstInterface^.stMultiCam.iq_stExt.xNoModuloMasterAtStart),
									q_etDiag	=> q_etDiag,
									q_etDiagExt	=> q_etDiagExt,
									q_sMsg		=> q_sMsg);

	IF q_etDiag <> GD.ET_Diag.Ok THEN
		RETURN;
	END_IF

	THIS^.fbTreeWriter.Parameter(	i_sName		:= 'xNoModuloSlaveAtStart',
									i_sValue	:= BOOL_TO_STRING(THIS^.pstInterface^.stMultiCam.iq_stExt.xNoModuloSlaveAtStart),
									q_etDiag	=> q_etDiag,
									q_etDiagExt	=> q_etDiagExt,
									q_sMsg		=> q_sMsg);

	IF q_etDiag <> GD.ET_Diag.Ok THEN
		RETURN;
	END_IF

	THIS^.fbTreeWriter.Parameter(	i_sName		:= 'xNoCyclicCams',
									i_sValue	:= BOOL_TO_STRING(THIS^.pstInterface^.stMultiCam.iq_stExt.xNoCyclicCams),
									q_etDiag	=> q_etDiag,
									q_etDiagExt	=> q_etDiagExt,
									q_sMsg		=> q_sMsg);

	IF q_etDiag <> GD.ET_Diag.Ok THEN
		RETURN;
	END_IF

	THIS^.fbTreeWriter.Parameter(	i_sName		:= 'xFirstCamNoXLimMin',
									i_sValue	:= BOOL_TO_STRING(THIS^.pstInterface^.stMultiCam.iq_stExt.xFirstCamNoXLimMin),
									q_etDiag	=> q_etDiag,
									q_etDiagExt	=> q_etDiagExt,
									q_sMsg		=> q_sMsg);

	IF q_etDiag <> GD.ET_Diag.Ok THEN
		RETURN;
	END_IF

	THIS^.fbTreeWriter.Parameter(	i_sName		:= 'xStopPositionSelect',
									i_sValue	:= BOOL_TO_STRING(THIS^.pstInterface^.stMultiCam.iq_stExt.xStopPositionSelect),
									q_etDiag	=> q_etDiag,
									q_etDiagExt	=> q_etDiagExt,
									q_sMsg		=> q_sMsg);

	IF q_etDiag <> GD.ET_Diag.Ok THEN
		RETURN;
	END_IF

	THIS^.fbTreeWriter.Parameter(	i_sName		:= 'lrStopPosition',
									i_sValue	:= LREAL_TO_STRING(THIS^.pstInterface^.stMultiCam.iq_stExt.lrStopPosition),
									q_etDiag	=> q_etDiag,
									q_etDiagExt	=> q_etDiagExt,
									q_sMsg		=> q_sMsg);

	IF q_etDiag <> GD.ET_Diag.Ok THEN
		RETURN;
	END_IF

	THIS^.fbTreeWriter.Parameter(	i_sName		:= 'lrStopVelocity',
									i_sValue	:= LREAL_TO_STRING(THIS^.pstInterface^.stMultiCam.iq_stExt.lrStopVelocity),
									q_etDiag	=> q_etDiag,
									q_etDiagExt	=> q_etDiagExt,
									q_sMsg		=> q_sMsg);

	IF q_etDiag <> GD.ET_Diag.Ok THEN
		RETURN;
	END_IF

	THIS^.fbTreeWriter.Parameter(	i_sName		:= 'lrStopAcceleration',
									i_sValue	:= LREAL_TO_STRING(THIS^.pstInterface^.stMultiCam.iq_stExt.lrStopAcceleration),
									q_etDiag	=> q_etDiag,
									q_etDiagExt	=> q_etDiagExt,
									q_sMsg		=> q_sMsg);

	IF q_etDiag <> GD.ET_Diag.Ok THEN
		RETURN;
	END_IF

	THIS^.fbTreeWriter.Parameter(	i_sName		:= 'lrStopDeceleration',
									i_sValue	:= LREAL_TO_STRING(THIS^.pstInterface^.stMultiCam.iq_stExt.lrStopDeceleration),
									q_etDiag	=> q_etDiag,
									q_etDiagExt	=> q_etDiagExt,
									q_sMsg		=> q_sMsg);

	IF q_etDiag <> GD.ET_Diag.Ok THEN
		RETURN;
	END_IF

	THIS^.fbTreeWriter.Parameter(	i_sName		:= 'lrStopJerk',
									i_sValue	:= LREAL_TO_STRING(THIS^.pstInterface^.stMultiCam.iq_stExt.lrStopJerk),
									q_etDiag	=> q_etDiag,
									q_etDiagExt	=> q_etDiagExt,
									q_sMsg		=> q_sMsg);

	IF q_etDiag <> GD.ET_Diag.Ok THEN
		RETURN;
	END_IF

	THIS^.fbTreeWriter.Parameter(	i_sName		:= 'xStartPositionSelect',
									i_sValue	:= BOOL_TO_STRING(THIS^.pstInterface^.stMultiCam.iq_stExt.xStartPositionSelect),
									q_etDiag	=> q_etDiag,
									q_etDiagExt	=> q_etDiagExt,
									q_sMsg		=> q_sMsg);

	IF q_etDiag <> GD.ET_Diag.Ok THEN
		RETURN;
	END_IF

	THIS^.fbTreeWriter.Parameter(	i_sName		:= 'lrStartPosition',
									i_sValue	:= LREAL_TO_STRING(THIS^.pstInterface^.stMultiCam.iq_stExt.lrStartPosition),
									q_etDiag	=> q_etDiag,
									q_etDiagExt	=> q_etDiagExt,
									q_sMsg		=> q_sMsg);

	IF q_etDiag <> GD.ET_Diag.Ok THEN
		RETURN;
	END_IF

	THIS^.fbTreeWriter.Parameter(	i_sName		:= 'lrStartVelocity',
									i_sValue	:= LREAL_TO_STRING(THIS^.pstInterface^.stMultiCam.iq_stExt.lrStartVelocity),
									q_etDiag	=> q_etDiag,
									q_etDiagExt	=> q_etDiagExt,
									q_sMsg		=> q_sMsg);

	IF q_etDiag <> GD.ET_Diag.Ok THEN
		RETURN;
	END_IF

	THIS^.fbTreeWriter.Parameter(	i_sName		:= 'lrStartAcceleration',
									i_sValue	:= LREAL_TO_STRING(THIS^.pstInterface^.stMultiCam.iq_stExt.lrStartAcceleration),
									q_etDiag	=> q_etDiag,
									q_etDiagExt	=> q_etDiagExt,
									q_sMsg		=> q_sMsg);

	IF q_etDiag <> GD.ET_Diag.Ok THEN
		RETURN;
	END_IF

	THIS^.fbTreeWriter.Parameter(	i_sName		:= 'lrStartDeceleration',
									i_sValue	:= LREAL_TO_STRING(THIS^.pstInterface^.stMultiCam.iq_stExt.lrStartDeceleration),
									q_etDiag	=> q_etDiag,
									q_etDiagExt	=> q_etDiagExt,
									q_sMsg		=> q_sMsg);

	IF q_etDiag <> GD.ET_Diag.Ok THEN
		RETURN;
	END_IF

	THIS^.fbTreeWriter.Parameter(	i_sName		:= 'lrStartJerk',
									i_sValue	:= LREAL_TO_STRING(THIS^.pstInterface^.stMultiCam.iq_stExt.lrStartJerk),
									q_etDiag	=> q_etDiag,
									q_etDiagExt	=> q_etDiagExt,
									q_sMsg		=> q_sMsg);

	IF q_etDiag <> GD.ET_Diag.Ok THEN
		RETURN;
	END_IF

	THIS^.fbTreeWriter.Parameter(	i_sName		:= 'xYEqualCheck',
									i_sValue	:= BOOL_TO_STRING(THIS^.pstInterface^.stMultiCam.iq_stExt.xYEqualCheck),
									q_etDiag	=> q_etDiag,
									q_etDiagExt	=> q_etDiagExt,
									q_sMsg		=> q_sMsg);

	IF q_etDiag <> GD.ET_Diag.Ok THEN
		RETURN;
	END_IF

	THIS^.fbTreeWriter.Parameter(	i_sName		:= 'lrYEqualCheckAccuracy',
									i_sValue	:= LREAL_TO_STRING(THIS^.pstInterface^.stMultiCam.iq_stExt.lrYEqualCheckAccuracy),
									q_etDiag	=> q_etDiag,
									q_etDiagExt	=> q_etDiagExt,
									q_sMsg		=> q_sMsg);

	IF q_etDiag <> GD.ET_Diag.Ok THEN
		RETURN;
	END_IF

	THIS^.fbTreeWriter.Parameter(	i_sName		:= 'xNewCamDirectAccept',
									i_sValue	:= BOOL_TO_STRING(THIS^.pstInterface^.stMultiCam.iq_stExt.xNewCamDirectAccept),
									q_etDiag	=> q_etDiag,
									q_etDiagExt	=> q_etDiagExt,
									q_sMsg		=> q_sMsg);

	IF q_etDiag <> GD.ET_Diag.Ok THEN
		RETURN;
	END_IF

	THIS^.fbTreeWriter.Parameter(	i_sName		:= 'xDisableLowEnd',
									i_sValue	:= BOOL_TO_STRING(THIS^.pstInterface^.stMultiCam.iq_stExt.xDisableLowEnd),
									q_etDiag	=> q_etDiag,
									q_etDiagExt	=> q_etDiagExt,
									q_sMsg		=> q_sMsg);

	IF q_etDiag <> GD.ET_Diag.Ok THEN
		RETURN;
	END_IF

	THIS^.fbTreeWriter.Parameter(	i_sName		:= 'xDisableHighEnd',
									i_sValue	:= BOOL_TO_STRING(THIS^.pstInterface^.stMultiCam.iq_stExt.xDisableHighEnd),
									q_etDiag	=> q_etDiag,
									q_etDiagExt	=> q_etDiagExt,
									q_sMsg		=> q_sMsg);

	IF q_etDiag <> GD.ET_Diag.Ok THEN
		RETURN;
	END_IF

	THIS^.fbTreeWriter.Parameter(	i_sName		:= 'lrCsMasterPosition',
									i_sValue	:= LREAL_TO_STRING(THIS^.pstInterface^.stMultiCam.iq_stExt.lrCsMasterPosition),
									q_etDiag	=> q_etDiag,
									q_etDiagExt	=> q_etDiagExt,
									q_sMsg		=> q_sMsg);

	IF q_etDiag <> GD.ET_Diag.Ok THEN
		RETURN;
	END_IF

	THIS^.fbTreeWriter.Parameter(	i_sName		:= 'xInWindowCheckWithoutLimits',
									i_sValue	:= BOOL_TO_STRING(THIS^.pstInterface^.stMultiCam.iq_stExt.xInWindowCheckWithoutLimits),
									q_etDiag	=> q_etDiag,
									q_etDiagExt	=> q_etDiagExt,
									q_sMsg		=> q_sMsg);

	IF q_etDiag <> GD.ET_Diag.Ok THEN
		RETURN;
	END_IF

	THIS^.fbTreeWriter.Parameter(	i_sName		:= 'etInWindowMode',
									i_sValue	:= AXM_FC_EtMultiCamWsModeToString(THIS^.pstInterface^.stMultiCam.iq_stExt.etInWindowMode),
									q_etDiag	=> q_etDiag,
									q_etDiagExt	=> q_etDiagExt,
									q_sMsg		=> q_sMsg);

	IF q_etDiag <> GD.ET_Diag.Ok THEN
		RETURN;
	END_IF

	THIS^.fbTreeWriter.Parameter(	i_sName		:= 'lrXStart',
									i_sValue	:= LREAL_TO_STRING(THIS^.pstInterface^.stMultiCam.iq_stExt.lrXStart),
									q_etDiag	=> q_etDiag,
									q_etDiagExt	=> q_etDiagExt,
									q_sMsg		=> q_sMsg);

	IF q_etDiag <> GD.ET_Diag.Ok THEN
		RETURN;
	END_IF

	THIS^.fbTreeWriter.Parameter(	i_sName		:= 'lrXIncr',
									i_sValue	:= LREAL_TO_STRING(THIS^.pstInterface^.stMultiCam.iq_stExt.lrXIncr),
									q_etDiag	=> q_etDiag,
									q_etDiagExt	=> q_etDiagExt,
									q_sMsg		=> q_sMsg);

	IF q_etDiag <> GD.ET_Diag.Ok THEN
		RETURN;
	END_IF

	THIS^.fbTreeWriter.Parameter(	i_sName		:= 'lrAccuracy',
									i_sValue	:= LREAL_TO_STRING(THIS^.pstInterface^.stMultiCam.iq_stExt.lrAccuracy),
									q_etDiag	=> q_etDiag,
									q_etDiagExt	=> q_etDiagExt,
									q_sMsg		=> q_sMsg);

	IF q_etDiag <> GD.ET_Diag.Ok THEN
		RETURN;
	END_IF

THIS^.fbTreeWriter.NodeEnd(	q_etDiag	=> q_etDiag,
							q_etDiagExt	=> q_etDiagExt,
							q_sMsg		=> q_sMsg);

IF q_etDiag <> GD.ET_Diag.Ok THEN
	RETURN;
END_IF

(* ---- WriteInterfaceMultiCamMotionParCamPoint.meth.st ---- *)
{attribute 'conditionalshow_all_locals'}
METHOD INTERNAL WriteInterfaceMultiCamMotionParCamPoint : BOOL
VAR_INPUT
END_VAR
VAR_OUTPUT
	q_etDiag		: GD.ET_Diag;
	q_etDiagExt	: TPL.ET_DiagExt;
	q_sMsg			: STRING[80];
END_VAR

THIS^.fbTreeWriter.NodeStart(	i_sName		:= Standard.CONCAT('astCamPoint[', Standard.CONCAT(DINT_TO_STRING(THIS^.diCamPointCounter), ']')),
								q_etDiag	=> q_etDiag,
								q_etDiagExt	=> q_etDiagExt,
								q_sMsg		=> q_sMsg);

IF q_etDiag <> GD.ET_Diag.Ok THEN
	RETURN;
END_IF

	THIS^.fbTreeWriter.Parameter(	i_sName		:= 'lrX',
									i_sValue	:= LREAL_TO_STRING(THIS^.pstInterface^.stMultiCam.iq_astMotionPar[THIS^.diMotionParCounter].astCamPoint[THIS^.diCamPointCounter].lrX),
									q_etDiag	=> q_etDiag,
									q_etDiagExt	=> q_etDiagExt,
									q_sMsg		=> q_sMsg);

	IF q_etDiag <> GD.ET_Diag.Ok THEN
		RETURN;
	END_IF

	THIS^.fbTreeWriter.Parameter(	i_sName		:= 'lrY',
									i_sValue	:= LREAL_TO_STRING(THIS^.pstInterface^.stMultiCam.iq_astMotionPar[THIS^.diMotionParCounter].astCamPoint[THIS^.diCamPointCounter].lrY),
									q_etDiag	=> q_etDiag,
									q_etDiagExt	=> q_etDiagExt,
									q_sMsg		=> q_sMsg);

	IF q_etDiag <> GD.ET_Diag.Ok THEN
		RETURN;
	END_IF

	THIS^.fbTreeWriter.Parameter(	i_sName		:= 'etCamType',
									i_sValue	:= AXM_FC_EtCamTypeToString(THIS^.pstInterface^.stMultiCam.iq_astMotionPar[THIS^.diMotionParCounter].astCamPoint[THIS^.diCamPointCounter].etCamType),
									q_etDiag	=> q_etDiag,
									q_etDiagExt	=> q_etDiagExt,
									q_sMsg		=> q_sMsg);

	IF q_etDiag <> GD.ET_Diag.Ok THEN
		RETURN;
	END_IF

	THIS^.fbTreeWriter.Parameter(	i_sName		:= 'lrM',
									i_sValue	:= LREAL_TO_STRING(THIS^.pstInterface^.stMultiCam.iq_astMotionPar[THIS^.diMotionParCounter].astCamPoint[THIS^.diCamPointCounter].lrM),
									q_etDiag	=> q_etDiag,
									q_etDiagExt	=> q_etDiagExt,
									q_sMsg		=> q_sMsg);

	IF q_etDiag <> GD.ET_Diag.Ok THEN
		RETURN;
	END_IF

	THIS^.fbTreeWriter.Parameter(	i_sName		:= 'lrK',
									i_sValue	:= LREAL_TO_STRING(THIS^.pstInterface^.stMultiCam.iq_astMotionPar[THIS^.diMotionParCounter].astCamPoint[THIS^.diCamPointCounter].lrK),
									q_etDiag	=> q_etDiag,
									q_etDiagExt	=> q_etDiagExt,
									q_sMsg		=> q_sMsg);

	IF q_etDiag <> GD.ET_Diag.Ok THEN
		RETURN;
	END_IF

	THIS^.fbTreeWriter.Parameter(	i_sName		:= 'lrYUser',
									i_sValue	:= LREAL_TO_STRING(THIS^.pstInterface^.stMultiCam.iq_astMotionPar[THIS^.diMotionParCounter].astCamPoint[THIS^.diCamPointCounter].lrYUser),
									q_etDiag	=> q_etDiag,
									q_etDiagExt	=> q_etDiagExt,
									q_sMsg		=> q_sMsg);

	IF q_etDiag <> GD.ET_Diag.Ok THEN
		RETURN;
	END_IF

	THIS^.fbTreeWriter.Parameter(	i_sName		:= 'diProfileId',
									i_sValue	:= DINT_TO_STRING(THIS^.pstInterface^.stMultiCam.iq_astMotionPar[THIS^.diMotionParCounter].astCamPoint[THIS^.diCamPointCounter].diProfileId),
									q_etDiag	=> q_etDiag,
									q_etDiagExt	=> q_etDiagExt,
									q_sMsg		=> q_sMsg);

	IF q_etDiag <> GD.ET_Diag.Ok THEN
		RETURN;
	END_IF

	THIS^.fbTreeWriter.Parameter(	i_sName		:= 'lrYUserOffset',
									i_sValue	:= LREAL_TO_STRING(THIS^.pstInterface^.stMultiCam.iq_astMotionPar[THIS^.diMotionParCounter].astCamPoint[THIS^.diCamPointCounter].lrYUserOffset),
									q_etDiag	=> q_etDiag,
									q_etDiagExt	=> q_etDiagExt,
									q_sMsg		=> q_sMsg);

	IF q_etDiag <> GD.ET_Diag.Ok THEN
		RETURN;
	END_IF

	THIS^.fbTreeWriter.Parameter(	i_sName		:= 'lrLambda',
									i_sValue	:= LREAL_TO_STRING(THIS^.pstInterface^.stMultiCam.iq_astMotionPar[THIS^.diMotionParCounter].astCamPoint[THIS^.diCamPointCounter].lrLambda),
									q_etDiag	=> q_etDiag,
									q_etDiagExt	=> q_etDiagExt,
									q_sMsg		=> q_sMsg);

	IF q_etDiag <> GD.ET_Diag.Ok THEN
		RETURN;
	END_IF

	THIS^.fbTreeWriter.Parameter(	i_sName		:= 'lrC',
									i_sValue	:= LREAL_TO_STRING(THIS^.pstInterface^.stMultiCam.iq_astMotionPar[THIS^.diMotionParCounter].astCamPoint[THIS^.diCamPointCounter].lrC),
									q_etDiag	=> q_etDiag,
									q_etDiagExt	=> q_etDiagExt,
									q_sMsg		=> q_sMsg);

	IF q_etDiag <> GD.ET_Diag.Ok THEN
		RETURN;
	END_IF

THIS^.fbTreeWriter.NodeEnd(	q_etDiag	=> q_etDiag,
							q_etDiagExt	=> q_etDiagExt,
							q_sMsg		=> q_sMsg);

IF q_etDiag <> GD.ET_Diag.Ok THEN
	RETURN;
END_IF

(* ---- WriteInterfaceMultiCamMotionParCamPointEnd.meth.st ---- *)
{attribute 'conditionalshow_all_locals'}
METHOD INTERNAL WriteInterfaceMultiCamMotionParCamPointEnd : BOOL
VAR_INPUT
END_VAR
VAR_OUTPUT
	q_etDiag		: GD.ET_Diag;
	q_etDiagExt	: TPL.ET_DiagExt;
	q_sMsg			: STRING[80];
END_VAR

THIS^.fbTreeWriter.NodeEnd(	q_etDiag	=> q_etDiag,
							q_etDiagExt	=> q_etDiagExt,
							q_sMsg		=> q_sMsg);

IF q_etDiag <> GD.ET_Diag.Ok THEN
	RETURN;
END_IF

(* ---- WriteInterfaceMultiCamMotionParCamPointStart.meth.st ---- *)
{attribute 'conditionalshow_all_locals'}
METHOD INTERNAL WriteInterfaceMultiCamMotionParCamPointStart : BOOL
VAR_INPUT
END_VAR
VAR_OUTPUT
	q_etDiag		: GD.ET_Diag;
	q_etDiagExt	: TPL.ET_DiagExt;
	q_sMsg			: STRING[80];
END_VAR

THIS^.fbTreeWriter.NodeStart(	i_sName		:= 'astCamPoint',
								q_etDiag	=> q_etDiag,
								q_etDiagExt	=> q_etDiagExt,
								q_sMsg		=> q_sMsg);

IF q_etDiag <> GD.ET_Diag.Ok THEN
	RETURN;
END_IF

(* ---- WriteInterfaceMultiCamMotionParCyclicEnd.meth.st ---- *)
{attribute 'conditionalshow_all_locals'}
METHOD INTERNAL WriteInterfaceMultiCamMotionParCyclicEnd : BOOL
VAR_INPUT
END_VAR
VAR_OUTPUT
	q_etDiag		: GD.ET_Diag;
	q_etDiagExt	: TPL.ET_DiagExt;
	q_sMsg			: STRING[80];
END_VAR

THIS^.fbTreeWriter.NodeEnd(	q_etDiag	=> q_etDiag,
							q_etDiagExt	=> q_etDiagExt,
							q_sMsg		=> q_sMsg);

IF q_etDiag <> GD.ET_Diag.Ok THEN
	RETURN;
END_IF

(* ---- WriteInterfaceMultiCamMotionParCyclicStart.meth.st ---- *)
{attribute 'conditionalshow_all_locals'}
METHOD INTERNAL WriteInterfaceMultiCamMotionParCyclicStart : BOOL
VAR_INPUT
END_VAR
VAR_OUTPUT
	q_etDiag		: GD.ET_Diag;
	q_etDiagExt	: TPL.ET_DiagExt;
	q_sMsg			: STRING[80];
END_VAR

THIS^.fbTreeWriter.NodeStart(	i_sName		:= Standard.CONCAT('iq_astMotionPar[', Standard.CONCAT(DINT_TO_STRING(THIS^.diMotionParCounter), ']')),
								q_etDiag	=> q_etDiag,
								q_etDiagExt	=> q_etDiagExt,
								q_sMsg		=> q_sMsg);

IF q_etDiag <> GD.ET_Diag.Ok THEN
	RETURN;
END_IF

	THIS^.fbTreeWriter.Parameter(	i_sName		:= 'diNumberOfCamPoints',
									i_sValue	:= DINT_TO_STRING(THIS^.pstInterface^.stMultiCam.iq_astMotionPar[THIS^.diMotionParCounter].diNumberOfCamPoints),
									q_etDiag	=> q_etDiag,
									q_etDiagExt	=> q_etDiagExt,
									q_sMsg		=> q_sMsg);

	IF q_etDiag <> GD.ET_Diag.Ok THEN
		RETURN;
	END_IF

	THIS^.fbTreeWriter.Parameter(	i_sName		:= 'diUserTableId',
									i_sValue	:= DINT_TO_STRING(THIS^.pstInterface^.stMultiCam.iq_astMotionPar[THIS^.diMotionParCounter].diUserTableId),
									q_etDiag	=> q_etDiag,
									q_etDiagExt	=> q_etDiagExt,
									q_sMsg		=> q_sMsg);

	IF q_etDiag <> GD.ET_Diag.Ok THEN
		RETURN;
	END_IF

	THIS^.fbTreeWriter.Parameter(	i_sName		:= 'lrYPeriod',
									i_sValue	:= LREAL_TO_STRING(THIS^.pstInterface^.stMultiCam.iq_astMotionPar[THIS^.diMotionParCounter].lrYPeriod),
									q_etDiag	=> q_etDiag,
									q_etDiagExt	=> q_etDiagExt,
									q_sMsg		=> q_sMsg);

	IF q_etDiag <> GD.ET_Diag.Ok THEN
		RETURN;
	END_IF

(* ---- WriteInterfaceMultiCamMotionParEnd.meth.st ---- *)
METHOD INTERNAL WriteInterfaceMultiCamMotionParEnd : BOOL
VAR_INPUT
END_VAR
VAR_OUTPUT
	q_etDiag		: GD.ET_Diag;
	q_etDiagExt	: TPL.ET_DiagExt;
	q_sMsg			: STRING[80];
END_VAR

THIS^.fbTreeWriter.NodeEnd(	q_etDiag	=> q_etDiag,
							q_etDiagExt	=> q_etDiagExt,
							q_sMsg		=> q_sMsg);

(* ---- WriteInterfaceMultiCamMotionParStart.meth.st ---- *)
METHOD INTERNAL WriteInterfaceMultiCamMotionParStart : BOOL
VAR_INPUT
END_VAR
VAR_OUTPUT
	q_etDiag		: GD.ET_Diag;
	q_etDiagExt	: TPL.ET_DiagExt;
	q_sMsg			: STRING[80];
END_VAR

THIS^.fbTreeWriter.NodeStart(	i_sName		:= 'iq_astMotionPar',
								q_etDiag	=> q_etDiag,
								q_etDiagExt	=> q_etDiagExt,
								q_sMsg		=> q_sMsg);

(* ---- WriteInterfaceMultiCamParamIn.meth.st ---- *)
METHOD INTERNAL WriteInterfaceMultiCamParamIn : BOOL
VAR_INPUT
END_VAR
VAR_OUTPUT
	q_etDiag		: GD.ET_Diag;
	q_etDiagExt	: TPL.ET_DiagExt;
	q_sMsg			: STRING[80];
END_VAR

THIS^.fbTreeWriter.Parameter(	i_sName		:= 'i_etCsModeSlave',
								i_sValue	:= AXM_FC_EtMultiCamCsModeSlaveToString(THIS^.pstInterface^.stMultiCam.i_etCsModeSlave),
								q_etDiag	=> q_etDiag,
								q_etDiagExt	=> q_etDiagExt,
								q_sMsg		=> q_sMsg);

IF q_etDiag <> GD.ET_Diag.Ok THEN
	RETURN;
END_IF

THIS^.fbTreeWriter.Parameter(	i_sName		:= 'i_etCsModeMaster',
								i_sValue	:= AXM_FC_EtMultiCamCsModeMasterToString(THIS^.pstInterface^.stMultiCam.i_etCsModeMaster),
								q_etDiag	=> q_etDiag,
								q_etDiagExt	=> q_etDiagExt,
								q_sMsg		=> q_sMsg);

IF q_etDiag <> GD.ET_Diag.Ok THEN
	RETURN;
END_IF

THIS^.fbTreeWriter.Parameter(	i_sName		:= 'i_etWsMode',
								i_sValue	:= AXM_FC_EtMultiCamWsModeToString(THIS^.pstInterface^.stMultiCam.i_etWsMode),
								q_etDiag	=> q_etDiag,
								q_etDiagExt	=> q_etDiagExt,
								q_sMsg		=> q_sMsg);

IF q_etDiag <> GD.ET_Diag.Ok THEN
	RETURN;
END_IF

THIS^.fbTreeWriter.Parameter(	i_sName		:= 'i_lrWsWindow',
								i_sValue	:= LREAL_TO_STRING(THIS^.pstInterface^.stMultiCam.i_lrWsWindow),
								q_etDiag	=> q_etDiag,
								q_etDiagExt	=> q_etDiagExt,
								q_sMsg		=> q_sMsg);

IF q_etDiag <> GD.ET_Diag.Ok THEN
	RETURN;
END_IF

THIS^.fbTreeWriter.Parameter(	i_sName		:= 'i_lrWsVel',
								i_sValue	:= LREAL_TO_STRING(THIS^.pstInterface^.stMultiCam.i_lrWsVel),
								q_etDiag	=> q_etDiag,
								q_etDiagExt	=> q_etDiagExt,
								q_sMsg		=> q_sMsg);

IF q_etDiag <> GD.ET_Diag.Ok THEN
	RETURN;
END_IF

THIS^.fbTreeWriter.Parameter(	i_sName		:= 'i_lrWsAcc',
								i_sValue	:= LREAL_TO_STRING(THIS^.pstInterface^.stMultiCam.i_lrWsAcc),
								q_etDiag	=> q_etDiag,
								q_etDiagExt	=> q_etDiagExt,
								q_sMsg		=> q_sMsg);

IF q_etDiag <> GD.ET_Diag.Ok THEN
	RETURN;
END_IF

THIS^.fbTreeWriter.Parameter(	i_sName		:= 'i_lrWsJerk',
								i_sValue	:= LREAL_TO_STRING(THIS^.pstInterface^.stMultiCam.i_lrWsJerk),
								q_etDiag	=> q_etDiag,
								q_etDiagExt	=> q_etDiagExt,
								q_sMsg		=> q_sMsg);

IF q_etDiag <> GD.ET_Diag.Ok THEN
	RETURN;
END_IF

THIS^.fbTreeWriter.Parameter(	i_sName		:= 'i_xCheckEncoderPeriod',
								i_sValue	:= BOOL_TO_STRING(THIS^.pstInterface^.stMultiCam.i_xCheckEncoderPeriod),
								q_etDiag	=> q_etDiag,
								q_etDiagExt	=> q_etDiagExt,
								q_sMsg		=> q_sMsg);

IF q_etDiag <> GD.ET_Diag.Ok THEN
	RETURN;
END_IF

THIS^.fbTreeWriter.Parameter(	i_sName		:= 'i_xSetEncoderPosition',
								i_sValue	:= BOOL_TO_STRING(THIS^.pstInterface^.stMultiCam.i_xSetEncoderPosition),
								q_etDiag	=> q_etDiag,
								q_etDiagExt	=> q_etDiagExt,
								q_sMsg		=> q_sMsg);

IF q_etDiag <> GD.ET_Diag.Ok THEN
	RETURN;
END_IF

THIS^.fbTreeWriter.Parameter(	i_sName		:= 'i_lrSetEncoderOffset',
								i_sValue	:= LREAL_TO_STRING(THIS^.pstInterface^.stMultiCam.i_lrSetEncoderOffset),
								q_etDiag	=> q_etDiag,
								q_etDiagExt	=> q_etDiagExt,
								q_sMsg		=> q_sMsg);

IF q_etDiag <> GD.ET_Diag.Ok THEN
	RETURN;
END_IF

THIS^.fbTreeWriter.Parameter(	i_sName		:= 'i_diTXend',
								i_sValue	:= DINT_TO_STRING(THIS^.pstInterface^.stMultiCam.i_diTXend),
								q_etDiag	=> q_etDiag,
								q_etDiagExt	=> q_etDiagExt,
								q_sMsg		=> q_sMsg);

IF q_etDiag <> GD.ET_Diag.Ok THEN
	RETURN;
END_IF

THIS^.fbTreeWriter.Parameter(	i_sName		:= 'i_lrInstantXLimMax',
								i_sValue	:= LREAL_TO_STRING(THIS^.pstInterface^.stMultiCam.i_lrInstantXLimMax),
								q_etDiag	=> q_etDiag,
								q_etDiagExt	=> q_etDiagExt,
								q_sMsg		=> q_sMsg);

IF q_etDiag <> GD.ET_Diag.Ok THEN
	RETURN;
END_IF

THIS^.fbTreeWriter.Parameter(	i_sName		:= 'i_xEnableTabHandler',
								i_sValue	:= BOOL_TO_STRING(THIS^.pstInterface^.stMultiCam.i_xEnableTabHandler),
								q_etDiag	=> q_etDiag,
								q_etDiagExt	=> q_etDiagExt,
								q_sMsg		=> q_sMsg);

IF q_etDiag <> GD.ET_Diag.Ok THEN
	RETURN;
END_IF

THIS^.fbTreeWriter.Parameter(	i_sName		:= 'i_udiTableSelectNr',
								i_sValue	:= UDINT_TO_STRING(THIS^.pstInterface^.stMultiCam.i_udiTableSelectNr),
								q_etDiag	=> q_etDiag,
								q_etDiagExt	=> q_etDiagExt,
								q_sMsg		=> q_sMsg);

IF q_etDiag <> GD.ET_Diag.Ok THEN
	RETURN;
END_IF
